// TwinCAT 3 PLC project HalfBROTTests
// Title: HalfBROTTests
// Company: BROT
// ProjectVersion: 0.1.0
// ProgramVersion: 3.1.4024.66
// libraries:
//   HalfBROT, * (BROT)
//   BROTLib, 0.26.0 (BROT)
//   Tc2_Math, * (Beckhoff Automation GmbH)
//   Tc2_MC2, * (Beckhoff Automation GmbH)
//   Tc2_Standard, * (Beckhoff Automation GmbH)
//   Tc2_System, * (Beckhoff Automation GmbH)
//   Tc2_Utilities, * (Beckhoff Automation GmbH)
//   Tc3_Module, * (Beckhoff Automation GmbH)
//   VisuElemEventTable, 1.0.3.0 (System)
//   TcUnit, * (www.tcunit.org)
// project tree:
//   / PlcTask.TcTTO
//   POUs/ F_Note.TcPOU, GVL_Diag.TcGVL, FB_NullComm.TcPOU, FB_TestBase.TcPOU, FB_HydraulicsRig.TcPOU, FB_CoverRig.TcPOU, FB_PendantRig.TcPOU, FB_FocusUnlockRig.TcPOU, FB_HydraulicsControl_Tests.TcPOU, FB_CoverControl_Tests.TcPOU, FB_PendantControl_Tests.TcPOU, FB_FocusUnlock_Tests.TcPOU, FB_BrakeCloseHold_Tests.TcPOU, F_FocusHoldOnStop_Tests.TcPOU, MAIN.TcPOU
// real-time tasks:
//   TASK PlcTask: cycle T#10ms, priority 20, ADS port 350

CONFIGURATION HalfBROTTests
    RESOURCE PLC ON TwinCAT3
        TASK PlcTask(INTERVAL := T#10ms, PRIORITY := 20);
        PROGRAM MAIN WITH PlcTask : MAIN;
    END_RESOURCE
END_CONFIGURATION

// ---- POUs/GVL_Diag.TcGVL
{attribute 'qualified_only'}
VAR_GLOBAL
	// the failed checks of the scenario tests (F_Note), one "test: message;" each. Run-Tests.ps1 prints it when a test failed:
	// TcUnit itself only writes the failure text to the ADS log, which CI cannot see.
	sFailures	: STRING(1000);
END_VAR

// ---- POUs/MAIN.TcPOU
PROGRAM MAIN
VAR
	// TcUnit finds every FB_TestSuite instance by itself; it is enough to declare them here.
	fbHydraulicsTests	: FB_HydraulicsControl_Tests;
	fbCoverTests		: FB_CoverControl_Tests;
	fbPendantTests		: FB_PendantControl_Tests;
	fbFocusUnlockTests	: FB_FocusUnlock_Tests;
	fbBrakeCloseHoldTests	: FB_BrakeCloseHold_Tests;	// MONETcommon#277
	fbFocusHoldOnStopTests	: F_FocusHoldOnStop_Tests;	// MONETcommon#278
END_VAR

TcUnit.RUN();

END_PROGRAM

// ---- POUs/FB_HydraulicsControl_Tests.TcPOU
// Characterisation tests of HalfBROT.FB_HydraulicsControl (HalfBROT#32 step 3) through the I/O structs and the command methods
// (#30, #31): start-up, the brake (pressure delay, clearing, pressure loss, CloseBrake, pump stop, azimuth limit), the manual
// brake re-arm of #31, and the latched errors that need no more than 13 s. They pin what the block does today, they are
// not a specification. Every test owns a rig (FB_HydraulicsRig, a plant behind the structs) and runs over many PLC cycles;
// the block timers run on the system time, so the tests take real time (the longest about 15 s). The suction and
// pressure watchdogs are shortened through tSuctionWatchdog and tPressureWatchdog.
FUNCTION_BLOCK FB_HydraulicsControl_Tests EXTENDS FB_TestBase
VAR
END_VAR

Idle_Everything_Off();
Enable_Runs_Pump();
Open_Brake_After_Pressure_Delay();
No_Clearing_Keeps_Brake_Closed();
Pressure_Loss_Closes_Brake_Auto_Reopens();
CloseBrake_Closes_And_Ends_Request();
Pump_Stop_Closes_Brake();
Azimuth_Limit_Closes_Brake();
Manual_Brake_Stays_Closed_After_Pressure_Loss();
Manual_Brake_Reopens_After_Switch_Off_On();
Manual_Switch_Off_Closes_Brake();
Manual_Brake_Stays_Closed_After_Pump_Restart();
Oil_Low_Is_Error_Until_Reset();
Hydraulics_Watchdog_Is_Error();
Suction_Without_Feedback_Is_Error();
Missing_Pressure_Is_Error();
Main_Pump_Without_Feedback_Is_Error();

// No request, healthy sensors: no pump, no brake, no error, no starter reset.
METHOD PRIVATE Idle_Everything_Off
VAR_INST
	rig		: FB_HydraulicsRig;
	nStep	: INT;
	bViol	: BOOL;
END_VAR
TEST('Idle_Everything_Off');
sCurrent := 'Idle_Everything_Off: ';
IF nStep >= 90 THEN
	RETURN;
END_IF
rig.Scan();
IF rig.nScans >= 5 THEN
	Check(NOT rig.stOut.bOilPumpEnable, 'no pump enable');
	Check(NOT rig.stOut.bOilSuctionEnable, 'no suction enable');
	Check(NOT rig.stOut.bBrakeAzEl, 'brake output off');
	Check(NOT rig.fb.bError, 'no error with healthy sensors');
	Check(rig.fb.PumpState = HalfBROT.E_PumpState.Off, 'pump state Off');
	Check(rig.fb.bBrakeClosed AND NOT rig.fb.bBrakeOpen, 'brake reported closed');
	Check(rig.fb.BrakeState = HalfBROT.E_BrakeState.Closed, 'brake state Closed');
	Check(NOT rig.stOut.bResetOilPump AND NOT rig.stOut.bResetSuctionPump, 'no starter reset');
		nStep := 99;
		TEST_FINISHED();
END_IF
END_METHOD

// Enable starts the pump; the plant reports it running with pressure; the brake is not opened by the pump start.
METHOD PRIVATE Enable_Runs_Pump
VAR_INST
	rig		: FB_HydraulicsRig;
	nStep	: INT;
	bViol	: BOOL;
END_VAR
TEST('Enable_Runs_Pump');
sCurrent := 'Enable_Runs_Pump: ';
IF nStep >= 90 THEN
	RETURN;
END_IF
rig.Scan();
CASE nStep OF
0:
	rig.SetEnable(TRUE);
	rig.StepStart();
	nStep := 10;
10:
	IF rig.nStepScans >= 6 THEN
		Check(rig.fb.Enable, 'Enable reads back');
		Check(rig.stOut.bOilPumpEnable, 'pump enable output');
		Check(rig.fb.PumpRunning AND rig.fb.OilPressureOK, 'pump running and pressure reported');
		Check(rig.fb.PumpState = HalfBROT.E_PumpState.Running, 'pump state Running');
		Check(NOT rig.fb.Error, 'no error');
		Check(NOT rig.stOut.bBrakeAzEl, 'the pump start does not open the brake');
		nStep := 99;
		TEST_FINISHED();
	END_IF
END_CASE
END_METHOD

// OpenBrake() each scan: the brake output comes about 3 s after the pressure, the report 1 s after the output.
METHOD PRIVATE Open_Brake_After_Pressure_Delay
VAR_INST
	rig		: FB_HydraulicsRig;
	nStep	: INT;
	bViol	: BOOL;
END_VAR
TEST('Open_Brake_After_Pressure_Delay');
sCurrent := 'Open_Brake_After_Pressure_Delay: ';
IF nStep >= 90 THEN
	RETURN;
END_IF
rig.Scan();
CASE nStep OF
0:
	rig.bClearing := TRUE;
	rig.bAuto := TRUE;
	rig.SetEnable(TRUE);
	rig.StepStart();
	nStep := 10;
10:
	IF rig.StepTime(T#1S) THEN
		Check(NOT rig.stOut.bBrakeAzEl, 'no brake output during the pressure delay');
		nStep := 20;
	END_IF
20:
	IF rig.stOut.bBrakeAzEl THEN
		Check(rig.StepTime(T#2S500MS) AND NOT rig.StepTime(T#4S), 'the brake output comes about 3 s after the start');
		Check(NOT rig.fb.bBrakeOpen, 'open is reported 1 s after the output, not with it');
		Check(rig.fb.BrakeState = HalfBROT.E_BrakeState.Opening, 'brake state Opening while the output is on and not reported');
		rig.StepStart();
		nStep := 30;
	ELSIF rig.StepTime(T#6S) THEN
		Check(FALSE, 'the brake output never came');
		nStep := 99;
		TEST_FINISHED();
	END_IF
30:
	IF rig.fb.bBrakeOpen THEN
		Check(rig.StepTime(T#800MS) AND NOT rig.StepTime(T#2S), 'open is reported about 1 s after the output');
		Check(rig.fb.BrakeOpen AND NOT rig.fb.bBrakeClosed, 'BrakeOpen property and bBrakeClosed agree');
		Check(rig.fb.BrakeState = HalfBROT.E_BrakeState.Open, 'brake state Open when reported');
		nStep := 99;
		TEST_FINISHED();
	ELSIF rig.StepTime(T#3S) THEN
		Check(FALSE, 'open was never reported');
		nStep := 99;
		TEST_FINISHED();
	END_IF
END_CASE
END_METHOD

// Without bBrakeClearing the brake is not opened although it is requested and the pressure is there.
METHOD PRIVATE No_Clearing_Keeps_Brake_Closed
VAR_INST
	rig		: FB_HydraulicsRig;
	nStep	: INT;
	bViol	: BOOL;
END_VAR
TEST('No_Clearing_Keeps_Brake_Closed');
sCurrent := 'No_Clearing_Keeps_Brake_Closed: ';
IF nStep >= 90 THEN
	RETURN;
END_IF
rig.Scan();
CASE nStep OF
0:
	rig.bClearing := FALSE;
	rig.bAuto := TRUE;
	rig.SetEnable(TRUE);
	rig.StepStart();
	nStep := 10;
10:
	bViol := bViol OR rig.stOut.bBrakeAzEl OR rig.fb.bBrakeOpen;
	IF rig.StepTime(T#4S) THEN
		Check(NOT bViol, 'the brake stays closed without the clearing');
		Check(rig.fb.PumpRunning AND rig.fb.OilPressureOK, 'pump running with pressure');
		nStep := 99;
		TEST_FINISHED();
	END_IF
END_CASE
END_METHOD

// Pressure loss closes the brake after the 2 s debounce; with the automatic request still there it opens again after the pressure delay.
METHOD PRIVATE Pressure_Loss_Closes_Brake_Auto_Reopens
VAR_INST
	rig		: FB_HydraulicsRig;
	nStep	: INT;
	bViol	: BOOL;
END_VAR
TEST('Pressure_Loss_Closes_Brake_Auto_Reopens');
sCurrent := 'Pressure_Loss_Closes_Brake_Auto_Reopens: ';
IF nStep >= 90 THEN
	RETURN;
END_IF
rig.Scan();
CASE nStep OF
0:
	rig.bClearing := TRUE;
	rig.bAuto := TRUE;
	rig.SetEnable(TRUE);
	rig.StepStart();
	nStep := 10;
10:
	IF rig.fb.bBrakeOpen THEN
		rig.bPressure := FALSE;
		rig.StepStart();
		nStep := 20;
	ELSIF rig.StepTime(T#8S) THEN
		Check(FALSE, 'the brake never opened');
		nStep := 99;
		TEST_FINISHED();
	END_IF
20:
	IF NOT rig.stOut.bBrakeAzEl THEN
		Check(rig.StepTime(T#1S500MS), 'the brake holds during the 2 s debounce');
		Check(NOT rig.fb.bBrakeOpen, 'closed is reported');
		Check(rig.stOut.bOilPumpEnable, 'the pump enable stays');
		rig.bPressure := TRUE;
		rig.StepStart();
		nStep := 30;
	ELSIF rig.StepTime(T#4S) THEN
		Check(FALSE, 'the brake did not close on the pressure loss');
		nStep := 99;
		TEST_FINISHED();
	END_IF
30:
	IF rig.stOut.bBrakeAzEl THEN
		Check(rig.StepTime(T#2S), 'the brake opens again only after the pressure delay');
		nStep := 99;
		TEST_FINISHED();
	ELSIF rig.StepTime(T#6S) THEN
		Check(FALSE, 'the automatic request did not open the brake again');
		nStep := 99;
		TEST_FINISHED();
	END_IF
END_CASE
END_METHOD

// CloseBrake() closes the brake at once and the request ends: no automatic re-open without OpenBrake().
METHOD PRIVATE CloseBrake_Closes_And_Ends_Request
VAR_INST
	rig		: FB_HydraulicsRig;
	nStep	: INT;
	bViol	: BOOL;
END_VAR
TEST('CloseBrake_Closes_And_Ends_Request');
sCurrent := 'CloseBrake_Closes_And_Ends_Request: ';
IF nStep >= 90 THEN
	RETURN;
END_IF
rig.Scan();
CASE nStep OF
0:
	rig.bClearing := TRUE;
	rig.bAuto := TRUE;
	rig.SetEnable(TRUE);
	rig.StepStart();
	nStep := 10;
10:
	IF rig.fb.bBrakeOpen THEN
		rig.bAuto := FALSE;
		rig.fb.CloseBrake();
		rig.StepStart();
		nStep := 20;
	ELSIF rig.StepTime(T#8S) THEN
		Check(FALSE, 'the brake never opened');
		nStep := 99;
		TEST_FINISHED();
	END_IF
20:
	IF NOT rig.stOut.bBrakeAzEl THEN
		Check(NOT rig.StepTime(T#300MS), 'the brake output drops at once');
		Check(NOT rig.fb.bBrakeOpen, 'closed is reported');
		Check(rig.fb.BrakeState = HalfBROT.E_BrakeState.Closed, 'brake state Closed after the close');
		rig.StepStart();
		nStep := 30;
	ELSIF rig.StepTime(T#1S) THEN
		Check(FALSE, 'CloseBrake() did not close the brake');
		nStep := 99;
		TEST_FINISHED();
	END_IF
30:
	bViol := bViol OR rig.stOut.bBrakeAzEl;
	IF rig.StepTime(T#4S) THEN
		Check(NOT bViol, 'the brake stays closed with the pressure there');
		nStep := 99;
		TEST_FINISHED();
	END_IF
END_CASE
END_METHOD

// ManualStopPump drops the pump enable; with the pump the brake closes.
METHOD PRIVATE Pump_Stop_Closes_Brake
VAR_INST
	rig		: FB_HydraulicsRig;
	nStep	: INT;
	bViol	: BOOL;
END_VAR
TEST('Pump_Stop_Closes_Brake');
sCurrent := 'Pump_Stop_Closes_Brake: ';
IF nStep >= 90 THEN
	RETURN;
END_IF
rig.Scan();
CASE nStep OF
0:
	rig.bClearing := TRUE;
	rig.bAuto := TRUE;
	rig.SetEnable(TRUE);
	rig.StepStart();
	nStep := 10;
10:
	IF rig.fb.bBrakeOpen THEN
		rig.bAuto := FALSE;
		rig.SetStopPump(TRUE);
		rig.StepStart();
		nStep := 20;
	ELSIF rig.StepTime(T#8S) THEN
		Check(FALSE, 'the brake never opened');
		nStep := 99;
		TEST_FINISHED();
	END_IF
20:
	IF NOT rig.stOut.bBrakeAzEl THEN
		Check(NOT rig.StepTime(T#300MS), 'the brake output drops with the pump');
		Check(NOT rig.stOut.bOilPumpEnable, 'pump enable off');
		Check(NOT rig.fb.bBrakeOpen, 'closed is reported');
		nStep := 99;
		TEST_FINISHED();
	ELSIF rig.StepTime(T#1S) THEN
		Check(FALSE, 'the pump stop did not close the brake');
		nStep := 99;
		TEST_FINISHED();
	END_IF
END_CASE
END_METHOD

// The azimuth limit switch closes the brake and holds it closed while it is active, although the request goes on.
METHOD PRIVATE Azimuth_Limit_Closes_Brake
VAR_INST
	rig		: FB_HydraulicsRig;
	nStep	: INT;
	bViol	: BOOL;
END_VAR
TEST('Azimuth_Limit_Closes_Brake');
sCurrent := 'Azimuth_Limit_Closes_Brake: ';
IF nStep >= 90 THEN
	RETURN;
END_IF
rig.Scan();
CASE nStep OF
0:
	rig.bClearing := TRUE;
	rig.bAuto := TRUE;
	rig.SetEnable(TRUE);
	rig.StepStart();
	nStep := 10;
10:
	IF rig.fb.bBrakeOpen THEN
		rig.bAzLimit := TRUE;
		rig.StepStart();
		nStep := 20;
	ELSIF rig.StepTime(T#8S) THEN
		Check(FALSE, 'the brake never opened');
		nStep := 99;
		TEST_FINISHED();
	END_IF
20:
	IF NOT rig.stOut.bBrakeAzEl THEN
		Check(NOT rig.StepTime(T#300MS), 'the brake output drops at once');
		rig.StepStart();
		nStep := 30;
	ELSIF rig.StepTime(T#1S) THEN
		Check(FALSE, 'the azimuth limit did not close the brake');
		nStep := 99;
		TEST_FINISHED();
	END_IF
30:
	bViol := bViol OR rig.stOut.bBrakeAzEl;
	IF rig.StepTime(T#4S) THEN
		Check(NOT bViol, 'the brake stays closed while the limit is active');
		nStep := 99;
		TEST_FINISHED();
	END_IF
END_CASE
END_METHOD

// #31: the cabinet switch opens the brake once; after a pressure loss it stays closed while the switch stays on, with the pressure back.
METHOD PRIVATE Manual_Brake_Stays_Closed_After_Pressure_Loss
VAR_INST
	rig		: FB_HydraulicsRig;
	nStep	: INT;
	bViol	: BOOL;
END_VAR
TEST('Manual_Brake_Stays_Closed_After_Pressure_Loss');
sCurrent := 'Manual_Brake_Stays_Closed_After_Pressure_Loss: ';
IF nStep >= 90 THEN
	RETURN;
END_IF
rig.Scan();
CASE nStep OF
0:
	// the pump runs first: a switch edge before the pump runs is dropped by the block (the request is cleared while the pump is off)
	rig.bManual := TRUE;
	rig.SetEnable(TRUE);
	rig.StepStart();
	nStep := 5;
5:
	IF rig.StepTime(T#500MS) THEN
		rig.bSwitch := TRUE;
		rig.StepStart();
		nStep := 10;
	END_IF
10:
	IF rig.fb.bBrakeOpen THEN
		Check(rig.stOut.bBrakeAzEl, 'the switch opened the brake');
		rig.bPressure := FALSE;
		rig.StepStart();
		nStep := 20;
	ELSIF rig.StepTime(T#8S) THEN
		Check(FALSE, 'the brake never opened');
		nStep := 99;
		TEST_FINISHED();
	END_IF
20:
	IF NOT rig.stOut.bBrakeAzEl THEN
		Check(rig.StepTime(T#1S500MS), 'the brake holds during the 2 s debounce');
		rig.bPressure := TRUE;
		bViol := FALSE;
		rig.StepStart();
		nStep := 30;
	ELSIF rig.StepTime(T#4S) THEN
		Check(FALSE, 'the brake did not close on the pressure loss');
		nStep := 99;
		TEST_FINISHED();
	END_IF
30:
	bViol := bViol OR rig.stOut.bBrakeAzEl;
	IF rig.StepTime(T#4S500MS) THEN
		Check(rig.fb.bOilPressureOK AND rig.fb.PumpRunning, 'pressure is back');
		Check(NOT bViol, 'the brake is not opened again while the switch stays on');
		nStep := 99;
		TEST_FINISHED();
	END_IF
END_CASE
END_METHOD

// #31: after CloseBrake() the brake stays closed while the switch stays on; switch off and on opens it again.
METHOD PRIVATE Manual_Brake_Reopens_After_Switch_Off_On
VAR_INST
	rig		: FB_HydraulicsRig;
	nStep	: INT;
	bViol	: BOOL;
END_VAR
TEST('Manual_Brake_Reopens_After_Switch_Off_On');
sCurrent := 'Manual_Brake_Reopens_After_Switch_Off_On: ';
IF nStep >= 90 THEN
	RETURN;
END_IF
rig.Scan();
CASE nStep OF
0:
	// the pump runs first: a switch edge before the pump runs is dropped by the block (the request is cleared while the pump is off)
	rig.bManual := TRUE;
	rig.SetEnable(TRUE);
	rig.StepStart();
	nStep := 5;
5:
	IF rig.StepTime(T#500MS) THEN
		rig.bSwitch := TRUE;
		rig.StepStart();
		nStep := 10;
	END_IF
10:
	IF rig.fb.bBrakeOpen THEN
		rig.fb.CloseBrake();
		rig.StepStart();
		nStep := 20;
	ELSIF rig.StepTime(T#8S) THEN
		Check(FALSE, 'the brake never opened');
		nStep := 99;
		TEST_FINISHED();
	END_IF
20:
	IF NOT rig.stOut.bBrakeAzEl THEN
		Check(NOT rig.StepTime(T#300MS), 'CloseBrake() closes at once');
		bViol := FALSE;
		rig.StepStart();
		nStep := 30;
	ELSIF rig.StepTime(T#1S) THEN
		Check(FALSE, 'CloseBrake() did not close the brake');
		nStep := 99;
		TEST_FINISHED();
	END_IF
30:
	bViol := bViol OR rig.stOut.bBrakeAzEl;
	IF rig.StepTime(T#4S) THEN
		Check(NOT bViol, 'the brake stays closed while the switch stays on');
		rig.bSwitch := FALSE;
		rig.StepStart();
		nStep := 40;
	END_IF
40:
	IF rig.StepTime(T#500MS) THEN
		Check(NOT rig.stOut.bBrakeAzEl, 'the brake is closed with the switch off');
		rig.bSwitch := TRUE;
		rig.StepStart();
		nStep := 50;
	END_IF
50:
	IF rig.stOut.bBrakeAzEl THEN
		Check(NOT rig.StepTime(T#1S), 'the switch off and on opens the brake at once, the pressure delay has long run out');
		nStep := 99;
		TEST_FINISHED();
	ELSIF rig.StepTime(T#6S) THEN
		Check(FALSE, 'the brake did not open again after the switch went off and on');
		nStep := 99;
		TEST_FINISHED();
	END_IF
END_CASE
END_METHOD

// The permission: switch off closes the brake at once (bBrakeClearing) and ends the request.
METHOD PRIVATE Manual_Switch_Off_Closes_Brake
VAR_INST
	rig		: FB_HydraulicsRig;
	nStep	: INT;
	bViol	: BOOL;
END_VAR
TEST('Manual_Switch_Off_Closes_Brake');
sCurrent := 'Manual_Switch_Off_Closes_Brake: ';
IF nStep >= 90 THEN
	RETURN;
END_IF
rig.Scan();
CASE nStep OF
0:
	// the pump runs first: a switch edge before the pump runs is dropped by the block (the request is cleared while the pump is off)
	rig.bManual := TRUE;
	rig.SetEnable(TRUE);
	rig.StepStart();
	nStep := 5;
5:
	IF rig.StepTime(T#500MS) THEN
		rig.bSwitch := TRUE;
		rig.StepStart();
		nStep := 10;
	END_IF
10:
	IF rig.fb.bBrakeOpen THEN
		rig.bSwitch := FALSE;
		rig.StepStart();
		nStep := 20;
	ELSIF rig.StepTime(T#8S) THEN
		Check(FALSE, 'the brake never opened');
		nStep := 99;
		TEST_FINISHED();
	END_IF
20:
	IF NOT rig.stOut.bBrakeAzEl THEN
		Check(NOT rig.StepTime(T#300MS), 'the brake output drops at once');
		Check(NOT rig.fb.bBrakeOpen, 'closed is reported');
		Check(rig.fb.BrakeState = HalfBROT.E_BrakeState.Closed, 'brake state Closed after the close');
		nStep := 99;
		TEST_FINISHED();
	ELSIF rig.StepTime(T#1S) THEN
		Check(FALSE, 'the switch off did not close the brake');
		nStep := 99;
		TEST_FINISHED();
	END_IF
END_CASE
END_METHOD

// #31: a pump stop closes the brake; the pump runs again with the switch still on: the brake stays closed.
METHOD PRIVATE Manual_Brake_Stays_Closed_After_Pump_Restart
VAR_INST
	rig		: FB_HydraulicsRig;
	nStep	: INT;
	bViol	: BOOL;
END_VAR
TEST('Manual_Brake_Stays_Closed_After_Pump_Restart');
sCurrent := 'Manual_Brake_Stays_Closed_After_Pump_Restart: ';
IF nStep >= 90 THEN
	RETURN;
END_IF
rig.Scan();
CASE nStep OF
0:
	// the pump runs first: a switch edge before the pump runs is dropped by the block (the request is cleared while the pump is off)
	rig.bManual := TRUE;
	rig.SetEnable(TRUE);
	rig.StepStart();
	nStep := 5;
5:
	IF rig.StepTime(T#500MS) THEN
		rig.bSwitch := TRUE;
		rig.StepStart();
		nStep := 10;
	END_IF
10:
	IF rig.fb.bBrakeOpen THEN
		rig.SetStopPump(TRUE);
		rig.StepStart();
		nStep := 20;
	ELSIF rig.StepTime(T#8S) THEN
		Check(FALSE, 'the brake never opened');
		nStep := 99;
		TEST_FINISHED();
	END_IF
20:
	IF NOT rig.stOut.bBrakeAzEl THEN
		Check(NOT rig.StepTime(T#300MS), 'the pump stop closes the brake at once');
		rig.StepStart();
		nStep := 30;
	ELSIF rig.StepTime(T#1S) THEN
		Check(FALSE, 'the pump stop did not close the brake');
		nStep := 99;
		TEST_FINISHED();
	END_IF
30:
	IF rig.StepTime(T#500MS) THEN
		rig.SetStopPump(FALSE);
		bViol := FALSE;
		rig.StepStart();
		nStep := 40;
	END_IF
40:
	bViol := bViol OR rig.stOut.bBrakeAzEl;
	IF rig.StepTime(T#4S500MS) THEN
		Check(rig.fb.PumpRunning AND rig.fb.OilPressureOK, 'the pump runs again with pressure');
		Check(NOT bViol, 'the brake is not opened again while the switch stays on');
		nStep := 99;
		TEST_FINISHED();
	END_IF
END_CASE
END_METHOD

// Oil low is a latched error that stops the pump; Reset() clears it once the oil is back and the pump starts again (Enable is still set).
METHOD PRIVATE Oil_Low_Is_Error_Until_Reset
VAR_INST
	rig		: FB_HydraulicsRig;
	nStep	: INT;
	bViol	: BOOL;
END_VAR
TEST('Oil_Low_Is_Error_Until_Reset');
sCurrent := 'Oil_Low_Is_Error_Until_Reset: ';
IF nStep >= 90 THEN
	RETURN;
END_IF
rig.Scan();
CASE nStep OF
0:
	rig.SetEnable(TRUE);
	rig.StepStart();
	nStep := 10;
10:
	IF rig.nStepScans >= 5 THEN
		rig.stIn.bOilLow := FALSE;
		rig.StepStart();
		nStep := 20;
	END_IF
20:
	IF rig.nStepScans >= 3 THEN
		Check(rig.fb.Error AND rig.fb.bOilLow, 'oil low is an error');
		Check(rig.fb.PumpState = HalfBROT.E_PumpState.Error, 'pump state Error');
		Check(NOT rig.stOut.bOilPumpEnable, 'the error stops the pump');
		rig.stIn.bOilLow := TRUE;
		rig.StepStart();
		nStep := 30;
	END_IF
30:
	IF rig.nStepScans >= 3 THEN
		Check(rig.fb.Error, 'the error stays latched with the oil back');
		rig.fb.Reset();
		rig.StepStart();
		nStep := 40;
	END_IF
40:
	IF rig.nStepScans >= 4 THEN
		Check(NOT rig.fb.Error, 'Reset() clears the error');
		Check(rig.stOut.bOilPumpEnable, 'the pump starts again, Enable is still set');
		Check(rig.fb.PumpState = HalfBROT.E_PumpState.Running, 'pump state Running again after Reset()');
		nStep := 99;
		TEST_FINISHED();
	END_IF
END_CASE
END_METHOD

// The pump running without the suction pump for tHydraulicsWatchdog (1 s here, 140 s default, #10) is a latched error.
METHOD PRIVATE Hydraulics_Watchdog_Is_Error
VAR_INST
	rig		: FB_HydraulicsRig;
	nStep	: INT;
	bViol	: BOOL;
END_VAR
TEST('Hydraulics_Watchdog_Is_Error');
sCurrent := 'Hydraulics_Watchdog_Is_Error: ';
IF nStep >= 90 THEN
	RETURN;
END_IF
rig.Scan();
CASE nStep OF
0:
	rig.tHydraulicsWatchdog := T#1S;
	rig.bSuctionFollows := FALSE;
	rig.SetEnable(TRUE);
	rig.StepStart();
	nStep := 10;
10:
	bViol := bViol OR rig.fb.bHydraulicsFailure;
	IF rig.fb.Error THEN
		Check(rig.StepTime(T#800MS), 'not before the configured time');
		Check(bViol, 'the hydraulics failure was reported');
		Check(NOT rig.stOut.bOilPumpEnable, 'the error stops the pump');
		nStep := 99;
		TEST_FINISHED();
	ELSIF rig.StepTime(T#4S) THEN
		Check(FALSE, 'no hydraulics failure');
		nStep := 99;
		TEST_FINISHED();
	END_IF
END_CASE
END_METHOD

// The suction enable (manual start) without the run feedback for tSuctionWatchdog (1 s here, 15 s default) is a latched error.
METHOD PRIVATE Suction_Without_Feedback_Is_Error
VAR_INST
	rig		: FB_HydraulicsRig;
	nStep	: INT;
	bViol	: BOOL;
END_VAR
TEST('Suction_Without_Feedback_Is_Error');
sCurrent := 'Suction_Without_Feedback_Is_Error: ';
IF nStep >= 90 THEN
	RETURN;
END_IF
rig.Scan();
CASE nStep OF
0:
	rig.tSuctionWatchdog := T#1S;
	rig.bSuctionFollows := FALSE;
	rig.SetSuction(TRUE);
	rig.StepStart();
	nStep := 10;
10:
	bViol := bViol OR rig.fb.bSuctionFailure;
	IF rig.fb.Error THEN
		Check(rig.stOut.bOilSuctionEnable, 'the suction enable was on');
		Check(rig.StepTime(T#800MS), 'not before the configured time');
		Check(bViol, 'the suction failure was reported');
		nStep := 99;
		TEST_FINISHED();
	ELSIF rig.StepTime(T#4S) THEN
		Check(FALSE, 'no suction failure');
		nStep := 99;
		TEST_FINISHED();
	END_IF
END_CASE
END_METHOD

// The pump enabled without oil pressure for tPressureWatchdog (1 s here, 30 s default) is a latched error that stops the pump.
METHOD PRIVATE Missing_Pressure_Is_Error
VAR_INST
	rig		: FB_HydraulicsRig;
	nStep	: INT;
	bViol	: BOOL;
END_VAR
TEST('Missing_Pressure_Is_Error');
sCurrent := 'Missing_Pressure_Is_Error: ';
IF nStep >= 90 THEN
	RETURN;
END_IF
rig.Scan();
CASE nStep OF
0:
	rig.tPressureWatchdog := T#1S;
	rig.bPressure := FALSE;
	rig.SetEnable(TRUE);
	rig.StepStart();
	nStep := 10;
10:
	bViol := bViol OR rig.fb.bPressureFailure;
	IF rig.fb.Error THEN
		Check(rig.StepTime(T#800MS), 'not before the configured time');
		Check(bViol, 'the pressure failure was reported');
		Check(NOT rig.stOut.bOilPumpEnable, 'the error stops the pump');
		nStep := 99;
		TEST_FINISHED();
	ELSIF rig.StepTime(T#4S) THEN
		Check(FALSE, 'no pressure failure');
		nStep := 99;
		TEST_FINISHED();
	END_IF
END_CASE
END_METHOD

// No run feedback 10 s after the pump enable is a latched error (main pump failure).
METHOD PRIVATE Main_Pump_Without_Feedback_Is_Error
VAR_INST
	rig		: FB_HydraulicsRig;
	nStep	: INT;
	bViol	: BOOL;
END_VAR
TEST('Main_Pump_Without_Feedback_Is_Error');
sCurrent := 'Main_Pump_Without_Feedback_Is_Error: ';
IF nStep >= 90 THEN
	RETURN;
END_IF
rig.Scan();
CASE nStep OF
0:
	rig.bPumpFollows := FALSE;
	rig.SetEnable(TRUE);
	rig.StepStart();
	nStep := 10;
10:
	bViol := bViol OR rig.fb.bMainPumpFailure;
	IF rig.fb.Error THEN
		Check(rig.StepTime(T#9S500MS), 'not before the 10 s');
		Check(bViol, 'the main pump failure was reported');
		Check(NOT rig.stOut.bOilPumpEnable, 'the error stops the pump');
		nStep := 99;
		TEST_FINISHED();
	ELSIF rig.StepTime(T#13S) THEN
		Check(FALSE, 'no main pump failure');
		nStep := 99;
		TEST_FINISHED();
	END_IF
END_CASE
END_METHOD

END_FUNCTION_BLOCK

// ---- POUs/FB_TestBase.TcPOU
// Base of the HalfBROTTests suites: Check() is a TcUnit assertion that also notes a failed check in GVL_Diag.sFailures
// (printed by tools/Run-Tests.ps1, TcUnit itself writes the failure text only to the ADS log). The test method sets
// sCurrent to its name first.
FUNCTION_BLOCK FB_TestBase EXTENDS TcUnit.FB_TestSuite
VAR
	sCurrent	: STRING(80);
END_VAR

METHOD Check
VAR_INPUT
	bCondition	: BOOL;
	sMessage	: STRING(255);
END_VAR
AssertTrue(Condition := bCondition, Message := sMessage);
F_Note(bFailed := NOT bCondition, sText := CONCAT(sCurrent, sMessage));
END_METHOD

END_FUNCTION_BLOCK

// ---- POUs/F_Note.TcPOU
// Records a failed check in GVL_Diag.sFailures (see there). Called next to the TcUnit assertion, which does the actual test result.
FUNCTION F_Note : BOOL
VAR_INPUT
	bFailed	: BOOL;
	sText	: STRING(255);
END_VAR

IF bFailed AND LEN(GVL_Diag.sFailures) < 700 THEN
	GVL_Diag.sFailures := CONCAT(CONCAT(GVL_Diag.sFailures, sText), '; ');
END_IF
F_Note := bFailed;

END_FUNCTION

// ---- POUs/FB_HydraulicsRig.TcPOU
// FB_HydraulicsControl with a plant: the pump feedback follows the pump enable output one scan later and the oil pressure
// follows the pump (a starter and a pump that work), the suction feedback follows the suction enable. The sensors are healthy.
// bAuto calls OpenBrake() in every scan (the automatic request of MONETcommon), bManual calls ManualBrake(bSwitch) and
// feeds the switch to bBrakeClearing as MAIN of MONETS/MONETN does. tPumpResetPulse is T#0S: the pump starts at once.
// StepStart()/StepTime() measure real time from the start of a step (the block timers run on the system time).
FUNCTION_BLOCK FB_HydraulicsRig
VAR_INPUT
	stIn		: HalfBROT.ST_HydraulicsIn := (bOilLow := TRUE, bOilHigh := TRUE, bOilCold := TRUE, bOilFilterDirty := TRUE, nOilLevel := 8000);
	bClearing	: BOOL;
	bAzLimit	: BOOL;
	bAuto		: BOOL;
	bManual		: BOOL;
	bSwitch		: BOOL;
	bPumpFollows	: BOOL := TRUE;
	bPressure		: BOOL := TRUE;
	bSuctionFollows	: BOOL := TRUE;
	tHydraulicsWatchdog	: TIME := T#140S;
	tSuctionWatchdog	: TIME := T#15S;
	tPressureWatchdog	: TIME := T#30S;
END_VAR
VAR
	fbComm		: FB_NullComm;
	fb			: HalfBROT.FB_HydraulicsControl(comm := fbComm);
	stOut		: HalfBROT.ST_HydraulicsOut;
	tonStep		: TON;
	nScans		: UDINT;
	nStepScans	: UDINT;
END_VAR

METHOD Scan
nScans := nScans + 1;
nStepScans := nStepScans + 1;
IF bPumpFollows THEN
	stIn.bPumpRunning := stOut.bOilPumpEnable;
END_IF
stIn.bOilPressureOK := stIn.bPumpRunning AND bPressure;
IF bSuctionFollows THEN
	stIn.bSuctionRunning := stOut.bOilSuctionEnable;
END_IF
IF bAuto THEN
	fb.OpenBrake();
END_IF
IF bManual THEN
	bClearing := bSwitch;
	fb.ManualBrake(bSwitch := bSwitch);
END_IF
fb(stIn := stIn, bBrakeClearing := bClearing, bAzimuthLimitSwitch := bAzLimit, tHydraulicsWatchdog := tHydraulicsWatchdog,
	tSuctionWatchdog := tSuctionWatchdog, tPressureWatchdog := tPressureWatchdog, tPumpResetPulse := T#0S, stOut := stOut);
tonStep(IN := TRUE, PT := T#1H);
END_METHOD

METHOD StepStart
tonStep(IN := FALSE, PT := T#1H);
nStepScans := 0;
END_METHOD

METHOD StepTime : BOOL
VAR_INPUT
	tTime	: TIME;
END_VAR
StepTime := tonStep.ET >= tTime;
END_METHOD

METHOD SetEnable
VAR_INPUT
	bOn	: BOOL;
END_VAR
fb.Enable := bOn;
END_METHOD

METHOD SetSuction
VAR_INPUT
	bOn	: BOOL;
END_VAR
fb.ManualStartSuction := bOn;
END_METHOD

METHOD SetStopPump
VAR_INPUT
	bOn	: BOOL;
END_VAR
fb.ManualStopPump := bOn;
END_METHOD

END_FUNCTION_BLOCK

// ---- POUs/FB_NullComm.TcPOU
// Minimal I_Comm stub for tests: every Publish/PublishLog call is a no-op that reports success,
// so FBs under test can call fbComm.Publish(...) freely without a real MQTT connection.
FUNCTION_BLOCK FB_NullComm IMPLEMENTS BROTLib.I_Comm
VAR
END_VAR

METHOD Publish : BOOL
VAR_INPUT
	domain			: STRING(255) := 'environment';
	location		: STRING(255) := 'roof';
	parameter		: STRING(255);
	value			: STRING(255);
END_VAR
VAR_OUTPUT
	published	: BOOL;
END_VAR
Publish := TRUE;
published := TRUE;
END_METHOD

METHOD PublishLREAL : BOOL
VAR_INPUT
	domain			: STRING(255) := 'environment';
	location		: STRING(255) := 'roof';
	parameter		: STRING(255);
	value			: LREAL;
END_VAR
VAR_OUTPUT
	published	: BOOL;
END_VAR
PublishLREAL := TRUE;
published := TRUE;
END_METHOD

METHOD PublishINT : BOOL
VAR_INPUT
	domain			: STRING(255) := 'environment';
	location		: STRING(255) := 'roof';
	parameter		: STRING(255);
	value			: LINT;
END_VAR
VAR_OUTPUT
	published	: BOOL;
END_VAR
PublishINT := TRUE;
published := TRUE;
END_METHOD

METHOD PublishBOOL : BOOL
VAR_INPUT
	domain			: STRING(255) := 'environment';
	location		: STRING(255) := 'roof';
	parameter		: STRING(255);
	value			: BOOL;
END_VAR
VAR_OUTPUT
	published	: BOOL;
END_VAR
PublishBOOL := TRUE;
published := TRUE;
END_METHOD

METHOD PublishString : BOOL
VAR_INPUT
	domain			: STRING(255) := 'environment';
	location		: STRING(255) := 'roof';
	parameter		: STRING(255);
	value			: STRING(255);
END_VAR
VAR_OUTPUT
	published	: BOOL;
END_VAR
PublishString := TRUE;
published := TRUE;
END_METHOD

METHOD PublishLog : BOOL
VAR_INPUT
	level		: STRING(255) := 'INFO';
	message		: STRING(255);
END_VAR
VAR_OUTPUT
	published	: BOOL;
END_VAR
PublishLog := TRUE;
published := TRUE;
END_METHOD

END_FUNCTION_BLOCK

// ---- POUs/FB_CoverControl_Tests.TcPOU
// Characterisation tests of HalfBROT.FB_CoverControl (HalfBROT#32 step 3) through the I/O structs: the sequence 1->3->2 and
// 2->3->1, the last call of Open()/Close() wins, Stop(), the latched error of a limit switch fault (#28), the move timeout and
// the reversal dead time (#27). They pin what the block does today, they are not a specification. Every test owns a rig
// (FB_CoverRig, the limit switches set by hand) and runs over several PLC cycles; the timeout and reversal tests take real time.
FUNCTION_BLOCK FB_CoverControl_Tests EXTENDS FB_TestBase
VAR
END_VAR

Open_Sequence_1_3_2();
Close_Sequence_2_3_1();
Last_Call_Wins_Open_After_Close();
Last_Call_Wins_Close_After_Open();
Stop_Drops_Outputs_And_Command();
Limit_Switch_Fault_Stops_All_Until_Reset();
Move_Timeout_Is_Error();
Reversal_Waits_Dead_Time();

// Open(): cover 1 starts, cover 3 only when 1 is at its open switch, cover 2 only when 1 and 3 are; then all outputs are off.
METHOD PRIVATE Open_Sequence_1_3_2
VAR_INST
	rig		: FB_CoverRig;
	nStep	: INT;
	bViol	: BOOL;
END_VAR
TEST('Open_Sequence_1_3_2');
sCurrent := 'Open_Sequence_1_3_2: ';
IF nStep >= 90 THEN
	RETURN;
END_IF
rig.Scan();
CASE nStep OF
0:
	Check(rig.OpenOutputs() = '---' AND rig.CloseOutputs() = '---', CONCAT('no output without a command ', rig.State()));
	rig.fb.Open();
	nStep := 10;
10:
	Check(rig.OpenOutputs() = 'x--' AND rig.CloseOutputs() = '---', CONCAT('only cover 1 starts ', rig.State()));
	Check(rig.fb.State = HalfBROT.E_CoverState.Opening, CONCAT('state Opening ', rig.State()));
	rig.SetMid(1);
	nStep := 15;
15:
	Check(rig.OpenOutputs() = 'x--', CONCAT('cover 3 waits while cover 1 is on its way ', rig.State()));
	rig.SetOpen(1);
	nStep := 20;
20:
	Check(rig.OpenOutputs() = '--x', CONCAT('cover 3 starts when cover 1 is open ', rig.State()));
	rig.SetMid(3);
	nStep := 25;
25:
	Check(rig.OpenOutputs() = '--x', CONCAT('cover 2 waits while cover 3 is on its way ', rig.State()));
	rig.SetOpen(3);
	nStep := 30;
30:
	Check(rig.OpenOutputs() = '-x-', CONCAT('cover 2 starts when 1 and 3 are open ', rig.State()));
	rig.SetOpen(2);
	nStep := 40;
40:
	Check(rig.fb.bAllOpen AND rig.fb.Opened AND NOT rig.fb.Closed, CONCAT('all covers open ', rig.State()));
	Check(rig.fb.State = HalfBROT.E_CoverState.Idle, CONCAT('state Idle after the last cover ', rig.State()));
	Check(rig.OpenOutputs() = '---' AND rig.CloseOutputs() = '---', CONCAT('all outputs off ', rig.State()));
	nStep := 50;
50:
	Check(rig.OpenOutputs() = '---', CONCAT('the command ended with the last cover ', rig.State()));
	nStep := 99;
	TEST_FINISHED();
END_CASE
END_METHOD

// Close(): cover 2 starts, cover 3 only when 2 is at its closed switch, cover 1 only when 2 and 3 are; then all outputs are off.
METHOD PRIVATE Close_Sequence_2_3_1
VAR_INST
	rig		: FB_CoverRig;
	nStep	: INT;
	bViol	: BOOL;
END_VAR
TEST('Close_Sequence_2_3_1');
sCurrent := 'Close_Sequence_2_3_1: ';
IF nStep >= 90 THEN
	RETURN;
END_IF
rig.Scan();
CASE nStep OF
0:
	rig.AllOpen();
	nStep := 5;
5:
	Check(rig.OpenOutputs() = '---' AND rig.CloseOutputs() = '---', CONCAT('no output without a command ', rig.State()));
	rig.fb.Close();
	nStep := 10;
10:
	Check(rig.CloseOutputs() = '-x-' AND rig.OpenOutputs() = '---', CONCAT('only cover 2 starts ', rig.State()));
	Check(rig.fb.State = HalfBROT.E_CoverState.Closing, CONCAT('state Closing ', rig.State()));
	rig.SetMid(2);
	nStep := 15;
15:
	Check(rig.CloseOutputs() = '-x-', CONCAT('cover 3 waits while cover 2 is on its way ', rig.State()));
	rig.SetClosed(2);
	nStep := 20;
20:
	Check(rig.CloseOutputs() = '--x', CONCAT('cover 3 starts when cover 2 is closed ', rig.State()));
	rig.SetMid(3);
	nStep := 25;
25:
	Check(rig.CloseOutputs() = '--x', CONCAT('cover 1 waits while cover 3 is on its way ', rig.State()));
	rig.SetClosed(3);
	nStep := 30;
30:
	Check(rig.CloseOutputs() = 'x--', CONCAT('cover 1 starts when 2 and 3 are closed ', rig.State()));
	rig.SetClosed(1);
	nStep := 40;
40:
	Check(rig.fb.bAllClosed AND rig.fb.Closed AND NOT rig.fb.Opened, CONCAT('all covers closed ', rig.State()));
	Check(rig.OpenOutputs() = '---' AND rig.CloseOutputs() = '---', CONCAT('all outputs off ', rig.State()));
	nStep := 50;
50:
	Check(rig.CloseOutputs() = '---', CONCAT('the command ended with the last cover ', rig.State()));
	nStep := 99;
	TEST_FINISHED();
END_CASE
END_METHOD

// Close() then Open() in one cycle: the open request wins (Open() drops the close request).
METHOD PRIVATE Last_Call_Wins_Open_After_Close
VAR_INST
	rig		: FB_CoverRig;
	nStep	: INT;
	bViol	: BOOL;
END_VAR
TEST('Last_Call_Wins_Open_After_Close');
sCurrent := 'Last_Call_Wins_Open_After_Close: ';
IF nStep >= 90 THEN
	RETURN;
END_IF
rig.Scan();
CASE nStep OF
0:
	rig.AllMid();
	rig.fb.Close();
	rig.fb.Open();
	nStep := 10;
10:
	Check(rig.CloseOutputs() = '---', CONCAT('no close output ', rig.State()));
	Check(rig.OpenOutputs() = 'x--', CONCAT('cover 1 opens ', rig.State()));
	nStep := 99;
	TEST_FINISHED();
END_CASE
END_METHOD

// Open() then Close() in one cycle: the close request wins (Close() drops the open request).
METHOD PRIVATE Last_Call_Wins_Close_After_Open
VAR_INST
	rig		: FB_CoverRig;
	nStep	: INT;
	bViol	: BOOL;
END_VAR
TEST('Last_Call_Wins_Close_After_Open');
sCurrent := 'Last_Call_Wins_Close_After_Open: ';
IF nStep >= 90 THEN
	RETURN;
END_IF
rig.Scan();
CASE nStep OF
0:
	rig.AllMid();
	rig.fb.Open();
	rig.fb.Close();
	nStep := 10;
10:
	Check(rig.OpenOutputs() = '---', CONCAT('no open output ', rig.State()));
	Check(rig.CloseOutputs() = '-x-', CONCAT('cover 2 closes ', rig.State()));
	nStep := 99;
	TEST_FINISHED();
END_CASE
END_METHOD

// Stop() drops the running output in the next scan and the command with it: nothing restarts.
METHOD PRIVATE Stop_Drops_Outputs_And_Command
VAR_INST
	rig		: FB_CoverRig;
	nStep	: INT;
	bViol	: BOOL;
END_VAR
TEST('Stop_Drops_Outputs_And_Command');
sCurrent := 'Stop_Drops_Outputs_And_Command: ';
IF nStep >= 90 THEN
	RETURN;
END_IF
rig.Scan();
CASE nStep OF
0:
	rig.fb.Open();
	nStep := 10;
10:
	Check(rig.OpenOutputs() = 'x--', CONCAT('cover 1 opens ', rig.State()));
	rig.fb.Stop();
	nStep := 20;
20:
	Check(rig.OpenOutputs() = '---' AND rig.CloseOutputs() = '---', CONCAT('the outputs are off after Stop() ', rig.State()));
	nStep := 30;
30:
	Check(rig.OpenOutputs() = '---', CONCAT('nothing restarts ', rig.State()));
	nStep := 40;
40:
	Check(rig.OpenOutputs() = '---' AND NOT rig.fb.Error, CONCAT('still off, no error ', rig.State()));
	nStep := 99;
	TEST_FINISHED();
END_CASE
END_METHOD

// Both switches of one cover (#28): the error stops all covers and drops the command; it stays latched until Reset(), and the move needs a new Open() after it.
METHOD PRIVATE Limit_Switch_Fault_Stops_All_Until_Reset
VAR_INST
	rig		: FB_CoverRig;
	nStep	: INT;
	bViol	: BOOL;
END_VAR
TEST('Limit_Switch_Fault_Stops_All_Until_Reset');
sCurrent := 'Limit_Switch_Fault_Stops_All_Until_Reset: ';
IF nStep >= 90 THEN
	RETURN;
END_IF
rig.Scan();
CASE nStep OF
0:
	rig.fb.Open();
	nStep := 10;
10:
	Check(rig.OpenOutputs() = 'x--', CONCAT('cover 1 opens ', rig.State()));
	rig.SetBoth(3);
	nStep := 20;
20:
	Check(rig.fb.Error AND rig.fb.bError, CONCAT('the fault is an error ', rig.State()));
	Check(rig.fb.State = HalfBROT.E_CoverState.Error, CONCAT('state Error ', rig.State()));
	Check(rig.OpenOutputs() = '---' AND rig.CloseOutputs() = '---', CONCAT('all covers stop, also those without the fault ', rig.State()));
	rig.SetClosed(3);
	rig.fb.Open();
	nStep := 30;
30:
	Check(rig.fb.Error, CONCAT('the error stays latched with the switch fixed ', rig.State()));
	Check(rig.fb.State = HalfBROT.E_CoverState.Error, CONCAT('state stays Error until Reset() ', rig.State()));
	Check(rig.OpenOutputs() = '---', CONCAT('no output while the error is latched ', rig.State()));
	rig.fb.Reset();
	nStep := 40;
40:
	Check(NOT rig.fb.Error, CONCAT('Reset() clears the error ', rig.State()));
	Check(rig.fb.State = HalfBROT.E_CoverState.Idle, CONCAT('state Idle after Reset() ', rig.State()));
	Check(rig.OpenOutputs() = '---', CONCAT('the command was dropped by the error: nothing moves ', rig.State()));
	rig.fb.Open();
	nStep := 50;
50:
	Check(rig.OpenOutputs() = 'x--', CONCAT('a new Open() moves again ', rig.State()));
	nStep := 99;
	TEST_FINISHED();
END_CASE
END_METHOD

// A cover driven for tMoveTimeout (300 ms here, 60 s default) without reaching its switch stops and latches an error until Reset().
METHOD PRIVATE Move_Timeout_Is_Error
VAR_INST
	rig		: FB_CoverRig;
	nStep	: INT;
	bViol	: BOOL;
END_VAR
TEST('Move_Timeout_Is_Error');
sCurrent := 'Move_Timeout_Is_Error: ';
IF nStep >= 90 THEN
	RETURN;
END_IF
rig.Scan();
CASE nStep OF
0:
	rig.tMoveTimeout := T#300MS;
	rig.fb.Open();
	rig.StepStart();
	nStep := 10;
10:
	IF rig.fb.Error THEN
		Check(rig.StepTime(T#250MS), CONCAT('not before the timeout ', rig.State()));
		Check(rig.OpenOutputs() = '---', CONCAT('the output is off ', rig.State()));
		Check(rig.fb.State = HalfBROT.E_CoverState.Error, CONCAT('state Error after the timeout ', rig.State()));
		rig.fb.Reset();
		nStep := 20;
	ELSIF rig.StepTime(T#2S) THEN
		Check(FALSE, 'no timeout error');
		nStep := 99;
		TEST_FINISHED();
	END_IF
20:
	Check(NOT rig.fb.Error, CONCAT('Reset() clears the timeout error ', rig.State()));
	Check(rig.OpenOutputs() = '---', CONCAT('nothing moves by itself after the reset ', rig.State()));
	nStep := 99;
	TEST_FINISHED();
END_CASE
END_METHOD

// Open() under way, then Close() (#27): the close output waits tReversalDeadTime (300 ms here, 1 s default) after the open output dropped.
METHOD PRIVATE Reversal_Waits_Dead_Time
VAR_INST
	rig		: FB_CoverRig;
	nStep	: INT;
	bViol	: BOOL;
END_VAR
TEST('Reversal_Waits_Dead_Time');
sCurrent := 'Reversal_Waits_Dead_Time: ';
IF nStep >= 90 THEN
	RETURN;
END_IF
rig.Scan();
CASE nStep OF
0:
	rig.tReversalDeadTime := T#300MS;
	rig.fb.Open();
	nStep := 10;
10:
	Check(rig.OpenOutputs() = 'x--', CONCAT('cover 1 opens ', rig.State()));
	rig.SetMid(1);
	rig.fb.Close();
	rig.StepStart();
	nStep := 20;
20:
	Check(rig.OpenOutputs() = '---', CONCAT('the open output is dropped at once ', rig.State()));
	Check(rig.CloseOutputs() = '---', CONCAT('the close output waits for the dead time ', rig.State()));
	nStep := 30;
30:
	bViol := bViol OR (rig.CloseOutputs() <> '---' AND NOT rig.StepTime(T#250MS));
	IF rig.CloseOutputs() <> '---' THEN
		Check(NOT bViol, CONCAT('no close output before the dead time ', rig.State()));
		Check(rig.StepTime(T#250MS) AND NOT rig.StepTime(T#1S), CONCAT('the close output comes after the dead time ', rig.State()));
		Check(rig.CloseOutputs() = 'x--', CONCAT('cover 1 closes ', rig.State()));
		nStep := 99;
		TEST_FINISHED();
	ELSIF rig.StepTime(T#2S) THEN
		Check(FALSE, 'the close output never came');
		nStep := 99;
		TEST_FINISHED();
	END_IF
END_CASE
END_METHOD

END_FUNCTION_BLOCK

// ---- POUs/FB_CoverRig.TcPOU
// FB_CoverControl with limit switches the test sets by hand. The switches are inverted (TRUE = the cover is NOT at the
// switch), see the block: SetClosed(i) puts cover i at its closed switch, SetOpen(i) at its open switch, SetMid(i) between
// them, SetBoth(i) is the limit switch fault (both switches reached). All covers start closed.
// StepStart()/StepTime() measure real time from the start of a step (the block timers run on the system time).
FUNCTION_BLOCK FB_CoverRig
VAR_INPUT
	stIn		: HalfBROT.ST_CoverIn;
	tReversalDeadTime	: TIME := T#1S;
	tMoveTimeout		: TIME := T#60S;
END_VAR
VAR
	fbComm		: FB_NullComm;
	fb			: HalfBROT.FB_CoverControl(comm := fbComm);
	stOut		: HalfBROT.ST_CoverOut;
	tonStep		: TON;
	nScans		: UDINT;
	bInit		: BOOL;
	i			: INT;
END_VAR

METHOD Scan
IF NOT bInit THEN
	bInit := TRUE;
	FOR i := 1 TO 3 DO
		SetClosed(i);
	END_FOR
END_IF
nScans := nScans + 1;
fb(stIn := stIn, tReversalDeadTime := tReversalDeadTime, tMoveTimeout := tMoveTimeout, stOut := stOut);
tonStep(IN := TRUE, PT := T#1H);
END_METHOD

METHOD SetClosed
VAR_INPUT
	nCover	: INT;
END_VAR
stIn.abOpen[nCover] := TRUE;
stIn.abClosed[nCover] := FALSE;
END_METHOD

METHOD SetOpen
VAR_INPUT
	nCover	: INT;
END_VAR
stIn.abOpen[nCover] := FALSE;
stIn.abClosed[nCover] := TRUE;
END_METHOD

METHOD SetMid
VAR_INPUT
	nCover	: INT;
END_VAR
stIn.abOpen[nCover] := TRUE;
stIn.abClosed[nCover] := TRUE;
END_METHOD

METHOD SetBoth
VAR_INPUT
	nCover	: INT;
END_VAR
stIn.abOpen[nCover] := FALSE;
stIn.abClosed[nCover] := FALSE;
END_METHOD

METHOD AllOpen
FOR i := 1 TO 3 DO
	SetOpen(i);
END_FOR
END_METHOD

METHOD AllMid
FOR i := 1 TO 3 DO
	SetMid(i);
END_FOR
END_METHOD

METHOD OpenOutputs : STRING(3)
// the open outputs of cover 1, 2 and 3 as "x" or "-"
OpenOutputs := '';
FOR i := 1 TO 3 DO
	IF stOut.abOpen[i] THEN
		OpenOutputs := CONCAT(OpenOutputs, 'x');
	ELSE
		OpenOutputs := CONCAT(OpenOutputs, '-');
	END_IF
END_FOR
END_METHOD

METHOD CloseOutputs : STRING(3)
// the close outputs of cover 1, 2 and 3 as "x" or "-"
CloseOutputs := '';
FOR i := 1 TO 3 DO
	IF stOut.abClose[i] THEN
		CloseOutputs := CONCAT(CloseOutputs, 'x');
	ELSE
		CloseOutputs := CONCAT(CloseOutputs, '-');
	END_IF
END_FOR
END_METHOD

METHOD State : STRING(60)
State := CONCAT(CONCAT(CONCAT(CONCAT('[open ', OpenOutputs()), ' close '), CloseOutputs()), CONCAT(' err ', BOOL_TO_STRING(fb.bError)));
State := CONCAT(State, ']');
END_METHOD

METHOD StepStart
tonStep(IN := FALSE, PT := T#1H);
END_METHOD

METHOD StepTime : BOOL
VAR_INPUT
	tTime	: TIME;
END_VAR
StepTime := tonStep.ET >= tTime;
END_METHOD

END_FUNCTION_BLOCK

// ---- POUs/FB_PendantControl_Tests.TcPOU
// Characterisation tests of HalfBROT.FB_PendantControl (HalfBROT#32 step 3) through the I/O structs: the selector, the error
// lamp for selector 0 and for blocks that are not connected (#16), the covers (hold-to-run with the key on, the level with the
// key off, #5 cover part) and the hydraulics (start toggle, brake up/down). The focus, derotator, elevation, azimuth and
// telescope selections need their blocks and are only covered for "not connected". They pin what the block does today, they
// are not a specification. Every test owns a rig (FB_PendantRig, the pendant with the cover and hydraulics rigs behind it).
FUNCTION_BLOCK FB_PendantControl_Tests EXTENDS FB_TestBase
VAR
END_VAR

Selector_Decodes_BCD();
Selector_Zero_Lights_Error_Lamp_Only();
Selector_Without_Function_Has_No_Error();
Unset_References_Light_Error_Lamp();
Selector_14_Horn_And_Lamps_Follow_Key();
Cover_Lamps_Show_The_Switches();
Cover_Key_On_Hold_Up_Opens_Release_Stops();
Cover_Key_On_Hold_Down_Closes_Release_Stops();
Cover_Key_On_Up_And_Down_Together_Do_Nothing();
Cover_Run_Stops_When_Selector_Leaves_1_To_3();
Cover_Key_Off_Up_Opens();
Hydraulics_Start_Button_Toggles_Pump();
Hydraulics_Key_Off_Buttons_Do_Nothing();
Hydraulics_Up_Opens_Brake_Down_Closes();

// The four selector inputs are the bits 1, 2, 4 and 8 of Selection.
METHOD PRIVATE Selector_Decodes_BCD
VAR_INST
	rig		: FB_PendantRig;
	nStep	: INT;
	bViol	: BOOL;
END_VAR
TEST('Selector_Decodes_BCD');
sCurrent := 'Selector_Decodes_BCD: ';
IF nStep >= 90 THEN
	RETURN;
END_IF
rig.Scan();
CASE nStep OF
0:
	rig.SetSelector(1);
	rig.StepStart();
	nStep := 10;
10:
	IF rig.nStepScans >= 2 THEN
		Check(rig.fb.Selection = 1, CONCAT('selector 1 ', rig.State()));
		rig.SetSelector(2);
		rig.StepStart();
		nStep := 20;
	END_IF
20:
	IF rig.nStepScans >= 2 THEN
		Check(rig.fb.Selection = 2, CONCAT('selector 2 ', rig.State()));
		rig.SetSelector(4);
		rig.StepStart();
		nStep := 30;
	END_IF
30:
	IF rig.nStepScans >= 2 THEN
		Check(rig.fb.Selection = 4, CONCAT('selector 4 ', rig.State()));
		rig.SetSelector(8);
		rig.StepStart();
		nStep := 40;
	END_IF
40:
	IF rig.nStepScans >= 2 THEN
		Check(rig.fb.Selection = 8, CONCAT('selector 8 ', rig.State()));
		rig.SetSelector(11);
		rig.StepStart();
		nStep := 50;
	END_IF
50:
	IF rig.nStepScans >= 2 THEN
		Check(rig.fb.Selection = 11, CONCAT('selector 11 ', rig.State()));
		rig.SetSelector(15);
		rig.StepStart();
		nStep := 60;
	END_IF
60:
	IF rig.nStepScans >= 2 THEN
		Check(rig.fb.Selection = 15, CONCAT('selector 15 ', rig.State()));
		rig.SetSelector(0);
		rig.StepStart();
		nStep := 70;
	END_IF
70:
	IF rig.nStepScans >= 2 THEN
		Check(rig.fb.Selection = 0, CONCAT('selector 0 ', rig.State()));
		nStep := 99;
		TEST_FINISHED();
	END_IF
END_CASE
END_METHOD

// Selector at 0 (pendant disconnected): only the error lamp, whatever the buttons say; nothing moves (#12).
METHOD PRIVATE Selector_Zero_Lights_Error_Lamp_Only
VAR_INST
	rig		: FB_PendantRig;
	nStep	: INT;
	bViol	: BOOL;
END_VAR
TEST('Selector_Zero_Lights_Error_Lamp_Only');
sCurrent := 'Selector_Zero_Lights_Error_Lamp_Only: ';
IF nStep >= 90 THEN
	RETURN;
END_IF
rig.Scan();
CASE nStep OF
0:
	rig.SetSelector(0); rig.SetKey(TRUE); rig.SetUp(TRUE); rig.SetStart(TRUE);
	rig.StepStart();
	nStep := 10;
10:
	IF rig.nStepScans >= 6 THEN
		Check(rig.Lamps() = '----x', CONCAT('only the error lamp ', rig.State()));
		Check(rig.fb.State = HalfBROT.E_PendantState.Disconnected, CONCAT('state Disconnected ', rig.State()));
		Check(rig.cov.OpenOutputs() = '---' AND rig.cov.CloseOutputs() = '---', CONCAT('no cover moves ', rig.State()));
		Check(NOT rig.hyd.stOut.bOilPumpEnable, CONCAT('no pump ', rig.State()));
		nStep := 99;
		TEST_FINISHED();
	END_IF
END_CASE
END_METHOD

// Selector 4 (Nasmyth), 9 (dome) and 10 (filter wheel) do nothing and light no lamp, also with the key on.
METHOD PRIVATE Selector_Without_Function_Has_No_Error
VAR_INST
	rig		: FB_PendantRig;
	nStep	: INT;
	bViol	: BOOL;
END_VAR
TEST('Selector_Without_Function_Has_No_Error');
sCurrent := 'Selector_Without_Function_Has_No_Error: ';
IF nStep >= 90 THEN
	RETURN;
END_IF
rig.Scan();
CASE nStep OF
0:
	rig.SetKey(TRUE); rig.SetSelector(4);
	rig.StepStart();
	nStep := 10;
10:
	IF rig.nStepScans >= 3 THEN
		Check(rig.Lamps() = '-----', CONCAT('selector 4: no lamp ', rig.State()));
		rig.SetKey(TRUE); rig.SetSelector(9);
		rig.StepStart();
		nStep := 20;
	END_IF
20:
	IF rig.nStepScans >= 3 THEN
		Check(rig.Lamps() = '-----', CONCAT('selector 9: no lamp ', rig.State()));
		rig.SetKey(TRUE); rig.SetSelector(10);
		rig.StepStart();
		nStep := 30;
	END_IF
30:
	IF rig.nStepScans >= 3 THEN
		Check(rig.Lamps() = '-----', CONCAT('selector 10: no lamp ', rig.State()));
		nStep := 99;
		TEST_FINISHED();
	END_IF
END_CASE
END_METHOD

// Selections whose block is not connected (focus, derotator, elevation, azimuth, telescope) light the error lamp and do nothing, with key, start and up pressed: no access to the unset reference (#16).
METHOD PRIVATE Unset_References_Light_Error_Lamp
VAR_INST
	rig		: FB_PendantRig;
	nStep	: INT;
	bViol	: BOOL;
END_VAR
TEST('Unset_References_Light_Error_Lamp');
sCurrent := 'Unset_References_Light_Error_Lamp: ';
IF nStep >= 90 THEN
	RETURN;
END_IF
rig.Scan();
CASE nStep OF
0:
	rig.SetKey(TRUE); rig.SetStart(TRUE); rig.SetUp(TRUE); rig.SetSelector(5);
	rig.StepStart();
	nStep := 10;
10:
	IF rig.nStepScans >= 4 THEN
		Check(rig.Lamps() = '----x', CONCAT('selector 5: block not connected ', rig.State()));
		Check(rig.fb.State = HalfBROT.E_PendantState.ReferencesMissing, CONCAT('state ReferencesMissing ', rig.State()));
		rig.SetKey(TRUE); rig.SetStart(TRUE); rig.SetUp(TRUE); rig.SetSelector(6);
		rig.StepStart();
		nStep := 20;
	END_IF
20:
	IF rig.nStepScans >= 4 THEN
		Check(rig.Lamps() = '----x', CONCAT('selector 6: block not connected ', rig.State()));
		Check(rig.fb.State = HalfBROT.E_PendantState.ReferencesMissing, CONCAT('state ReferencesMissing ', rig.State()));
		rig.SetKey(TRUE); rig.SetStart(TRUE); rig.SetUp(TRUE); rig.SetSelector(7);
		rig.StepStart();
		nStep := 30;
	END_IF
30:
	IF rig.nStepScans >= 4 THEN
		Check(rig.Lamps() = '----x', CONCAT('selector 7: block not connected ', rig.State()));
		Check(rig.fb.State = HalfBROT.E_PendantState.ReferencesMissing, CONCAT('state ReferencesMissing ', rig.State()));
		rig.SetKey(TRUE); rig.SetStart(TRUE); rig.SetUp(TRUE); rig.SetSelector(8);
		rig.StepStart();
		nStep := 40;
	END_IF
40:
	IF rig.nStepScans >= 4 THEN
		Check(rig.Lamps() = '----x', CONCAT('selector 8: block not connected ', rig.State()));
		Check(rig.fb.State = HalfBROT.E_PendantState.ReferencesMissing, CONCAT('state ReferencesMissing ', rig.State()));
		rig.SetKey(TRUE); rig.SetStart(TRUE); rig.SetUp(TRUE); rig.SetSelector(11);
		rig.StepStart();
		nStep := 50;
	END_IF
50:
	IF rig.nStepScans >= 4 THEN
		Check(rig.Lamps() = '----x', CONCAT('selector 11: block not connected ', rig.State()));
		Check(rig.fb.State = HalfBROT.E_PendantState.ReferencesMissing, CONCAT('state ReferencesMissing ', rig.State()));
		rig.SetKey(TRUE); rig.SetStart(TRUE); rig.SetUp(TRUE); rig.SetSelector(12);
		rig.StepStart();
		nStep := 60;
	END_IF
60:
	IF rig.nStepScans >= 4 THEN
		Check(rig.Lamps() = '----x', CONCAT('selector 12: block not connected ', rig.State()));
		Check(rig.fb.State = HalfBROT.E_PendantState.ReferencesMissing, CONCAT('state ReferencesMissing ', rig.State()));
		rig.SetKey(TRUE); rig.SetStart(TRUE); rig.SetUp(TRUE); rig.SetSelector(13);
		rig.StepStart();
		nStep := 70;
	END_IF
70:
	IF rig.nStepScans >= 4 THEN
		Check(rig.Lamps() = '----x', CONCAT('selector 13: block not connected ', rig.State()));
		Check(rig.fb.State = HalfBROT.E_PendantState.ReferencesMissing, CONCAT('state ReferencesMissing ', rig.State()));
		nStep := 99;
		TEST_FINISHED();
	END_IF
END_CASE
END_METHOD

// Selector 14: lamps up, down, left and right and the horn follow the key switch.
METHOD PRIVATE Selector_14_Horn_And_Lamps_Follow_Key
VAR_INST
	rig		: FB_PendantRig;
	nStep	: INT;
	bViol	: BOOL;
END_VAR
TEST('Selector_14_Horn_And_Lamps_Follow_Key');
sCurrent := 'Selector_14_Horn_And_Lamps_Follow_Key: ';
IF nStep >= 90 THEN
	RETURN;
END_IF
rig.Scan();
CASE nStep OF
0:
	rig.SetSelector(14);
	rig.StepStart();
	nStep := 10;
10:
	IF rig.nStepScans >= 3 THEN
		Check(rig.Lamps() = '-----', CONCAT('key off: no lamp ', rig.State()));
		Check(rig.fb.State = HalfBROT.E_PendantState.Automatic, CONCAT('key off: state Automatic ', rig.State()));
		Check(NOT rig.fb.horn, CONCAT('key off: no horn ', rig.State()));
		rig.SetKey(TRUE);
		rig.StepStart();
		nStep := 20;
	END_IF
20:
	IF rig.nStepScans >= 3 THEN
		Check(rig.Lamps() = 'xxxx-', CONCAT('key on: four lamps, no error lamp ', rig.State()));
		Check(rig.fb.State = HalfBROT.E_PendantState.Manual, CONCAT('key on: state Manual ', rig.State()));
		Check(rig.fb.horn, CONCAT('key on: horn ', rig.State()));
		rig.SetKey(FALSE);
		rig.StepStart();
		nStep := 30;
	END_IF
30:
	IF rig.nStepScans >= 3 THEN
		Check(rig.Lamps() = '-----', CONCAT('key off again: no lamp ', rig.State()));
		Check(NOT rig.fb.horn, CONCAT('key off again: no horn ', rig.State()));
		nStep := 99;
		TEST_FINISHED();
	END_IF
END_CASE
END_METHOD

// Selector 1: up is lit while the cover is not at its open switch, down while it is not at its closed switch; with the key on the error lamp shows a limit switch fault.
METHOD PRIVATE Cover_Lamps_Show_The_Switches
VAR_INST
	rig		: FB_PendantRig;
	nStep	: INT;
	bViol	: BOOL;
END_VAR
TEST('Cover_Lamps_Show_The_Switches');
sCurrent := 'Cover_Lamps_Show_The_Switches: ';
IF nStep >= 90 THEN
	RETURN;
END_IF
rig.Scan();
CASE nStep OF
0:
	rig.SetSelector(1);
	rig.StepStart();
	nStep := 10;
10:
	IF rig.nStepScans >= 5 THEN
		Check(rig.Lamps() = 'x----', CONCAT('closed: up lit, down dark ', rig.State()));
		rig.cov.AllOpen();
		rig.StepStart();
		nStep := 20;
	END_IF
20:
	IF rig.nStepScans >= 5 THEN
		Check(rig.Lamps() = '-x---', CONCAT('open: up dark, down lit ', rig.State()));
		rig.cov.SetBoth(1); rig.SetKey(TRUE);
		rig.StepStart();
		nStep := 30;
	END_IF
30:
	IF rig.nStepScans >= 5 THEN
		Check(rig.Lamps() = '----x', CONCAT('both switches reached: error lamp ', rig.State()));
		rig.cov.SetMid(1);
		rig.StepStart();
		nStep := 40;
	END_IF
40:
	IF rig.nStepScans >= 5 THEN
		Check(rig.Lamps() = 'xx---', CONCAT('between the switches: up and down lit, no error ', rig.State()));
		nStep := 99;
		TEST_FINISHED();
	END_IF
END_CASE
END_METHOD

// Key on, selector 1: up held opens cover 1 (the block does the order); releasing the button stops the run.
METHOD PRIVATE Cover_Key_On_Hold_Up_Opens_Release_Stops
VAR_INST
	rig		: FB_PendantRig;
	nStep	: INT;
	bViol	: BOOL;
END_VAR
TEST('Cover_Key_On_Hold_Up_Opens_Release_Stops');
sCurrent := 'Cover_Key_On_Hold_Up_Opens_Release_Stops: ';
IF nStep >= 90 THEN
	RETURN;
END_IF
rig.Scan();
CASE nStep OF
0:
	rig.SetSelector(1); rig.SetKey(TRUE);
	rig.StepStart();
	nStep := 10;
10:
	IF rig.nStepScans >= 4 THEN
		Check(rig.cov.OpenOutputs() = '---' AND rig.cov.CloseOutputs() = '---', CONCAT('nothing moves without a button ', rig.State()));
		rig.SetUp(TRUE);
		rig.StepStart();
		nStep := 20;
	END_IF
20:
	IF rig.nStepScans >= 25 THEN
		Check(rig.cov.OpenOutputs() = 'x--' AND rig.cov.CloseOutputs() = '---', CONCAT('up held: cover 1 opens ', rig.State()));
		rig.SetUp(FALSE);
		rig.StepStart();
		nStep := 30;
	END_IF
30:
	IF rig.nStepScans >= 25 THEN
		Check(rig.cov.OpenOutputs() = '---' AND rig.cov.CloseOutputs() = '---', CONCAT('the release stops the run ', rig.State()));
		nStep := 99;
		TEST_FINISHED();
	END_IF
END_CASE
END_METHOD

// Key on, selector 1, all covers open: down held closes cover 2 first; releasing the button stops the run.
METHOD PRIVATE Cover_Key_On_Hold_Down_Closes_Release_Stops
VAR_INST
	rig		: FB_PendantRig;
	nStep	: INT;
	bViol	: BOOL;
END_VAR
TEST('Cover_Key_On_Hold_Down_Closes_Release_Stops');
sCurrent := 'Cover_Key_On_Hold_Down_Closes_Release_Stops: ';
IF nStep >= 90 THEN
	RETURN;
END_IF
rig.Scan();
CASE nStep OF
0:
	rig.cov.AllOpen(); rig.SetSelector(1); rig.SetKey(TRUE);
	rig.StepStart();
	nStep := 10;
10:
	IF rig.nStepScans >= 5 THEN
		Check(rig.cov.OpenOutputs() = '---' AND rig.cov.CloseOutputs() = '---', CONCAT('nothing moves without a button ', rig.State()));
		rig.SetDown(TRUE);
		rig.StepStart();
		nStep := 20;
	END_IF
20:
	IF rig.nStepScans >= 25 THEN
		Check(rig.cov.CloseOutputs() = '-x-' AND rig.cov.OpenOutputs() = '---', CONCAT('down held: cover 2 closes first ', rig.State()));
		rig.SetDown(FALSE);
		rig.StepStart();
		nStep := 30;
	END_IF
30:
	IF rig.nStepScans >= 5 THEN
		Check(rig.cov.OpenOutputs() = '---' AND rig.cov.CloseOutputs() = '---', CONCAT('the release stops the run ', rig.State()));
		nStep := 99;
		TEST_FINISHED();
	END_IF
END_CASE
END_METHOD

// Key on, selector 1: up and down pressed together start nothing.
METHOD PRIVATE Cover_Key_On_Up_And_Down_Together_Do_Nothing
VAR_INST
	rig		: FB_PendantRig;
	nStep	: INT;
	bViol	: BOOL;
END_VAR
TEST('Cover_Key_On_Up_And_Down_Together_Do_Nothing');
sCurrent := 'Cover_Key_On_Up_And_Down_Together_Do_Nothing: ';
IF nStep >= 90 THEN
	RETURN;
END_IF
rig.Scan();
CASE nStep OF
0:
	rig.SetSelector(1); rig.SetKey(TRUE); rig.SetUp(TRUE); rig.SetDown(TRUE);
	rig.StepStart();
	nStep := 10;
10:
	IF rig.nStepScans >= 12 THEN
		Check(rig.cov.OpenOutputs() = '---' AND rig.cov.CloseOutputs() = '---', CONCAT('up and down together ', rig.State()));
		nStep := 99;
		TEST_FINISHED();
	END_IF
END_CASE
END_METHOD

// A run started by the pendant stops when the selector leaves 1 to 3 although the button is still held.
METHOD PRIVATE Cover_Run_Stops_When_Selector_Leaves_1_To_3
VAR_INST
	rig		: FB_PendantRig;
	nStep	: INT;
	bViol	: BOOL;
END_VAR
TEST('Cover_Run_Stops_When_Selector_Leaves_1_To_3');
sCurrent := 'Cover_Run_Stops_When_Selector_Leaves_1_To_3: ';
IF nStep >= 90 THEN
	RETURN;
END_IF
rig.Scan();
CASE nStep OF
0:
	rig.SetSelector(1); rig.SetKey(TRUE); rig.SetUp(TRUE);
	rig.StepStart();
	nStep := 10;
10:
	IF rig.nStepScans >= 6 THEN
		Check(rig.cov.OpenOutputs() = 'x--', CONCAT('cover 1 opens ', rig.State()));
		rig.SetSelector(4);
		rig.StepStart();
		nStep := 20;
	END_IF
20:
	IF rig.nStepScans >= 4 THEN
		Check(rig.cov.OpenOutputs() = '---' AND rig.cov.CloseOutputs() = '---', CONCAT('the run stops with the selector ', rig.State()));
		nStep := 99;
		TEST_FINISHED();
	END_IF
END_CASE
END_METHOD

// Key off (automatic), selector 1: up opens cover 1 (the level, no hold-to-run).
METHOD PRIVATE Cover_Key_Off_Up_Opens
VAR_INST
	rig		: FB_PendantRig;
	nStep	: INT;
	bViol	: BOOL;
END_VAR
TEST('Cover_Key_Off_Up_Opens');
sCurrent := 'Cover_Key_Off_Up_Opens: ';
IF nStep >= 90 THEN
	RETURN;
END_IF
rig.Scan();
CASE nStep OF
0:
	rig.SetSelector(1); rig.SetUp(TRUE);
	rig.StepStart();
	nStep := 10;
10:
	IF rig.nStepScans >= 6 THEN
		Check(rig.cov.OpenOutputs() = 'x--' AND rig.cov.CloseOutputs() = '---', CONCAT('up: cover 1 opens ', rig.State()));
		nStep := 99;
		TEST_FINISHED();
	END_IF
END_CASE
END_METHOD

// Key on, selector 15: each press of start (the edge, not the level) toggles the hydraulics enable; the lamps show pump and pressure.
METHOD PRIVATE Hydraulics_Start_Button_Toggles_Pump
VAR_INST
	rig		: FB_PendantRig;
	nStep	: INT;
	bViol	: BOOL;
END_VAR
TEST('Hydraulics_Start_Button_Toggles_Pump');
sCurrent := 'Hydraulics_Start_Button_Toggles_Pump: ';
IF nStep >= 90 THEN
	RETURN;
END_IF
rig.Scan();
CASE nStep OF
0:
	rig.SetSelector(15); rig.SetKey(TRUE);
	rig.StepStart();
	nStep := 10;
10:
	IF rig.nStepScans >= 4 THEN
		Check(NOT rig.hyd.stOut.bOilPumpEnable, CONCAT('the pump is off ', rig.State()));
		rig.SetStart(TRUE);
		rig.StepStart();
		nStep := 20;
	END_IF
20:
	IF rig.nStepScans >= 15 THEN
		Check(rig.hyd.stOut.bOilPumpEnable AND rig.hyd.fb.Enable, CONCAT('the pump is enabled ', rig.State()));
		Check(rig.hyd.fb.PumpRunning AND rig.hyd.fb.OilPressureOK, CONCAT('pump running with pressure ', rig.State()));
		Check(rig.stOut.bLampLeft AND rig.stOut.bLampUp AND NOT rig.stOut.bLampDown, CONCAT('lamps: pump running, pressure, brake closed ', rig.State()));
		rig.SetStart(FALSE);
		rig.StepStart();
		nStep := 30;
	END_IF
30:
	IF rig.nStepScans >= 8 THEN
		Check(rig.hyd.stOut.bOilPumpEnable AND rig.hyd.fb.Enable, CONCAT('the pump is still enabled after the button was held and released ', rig.State()));
		rig.SetStart(TRUE);
		rig.StepStart();
		nStep := 40;
	END_IF
40:
	IF rig.nStepScans >= 8 THEN
		Check(NOT rig.hyd.stOut.bOilPumpEnable AND NOT rig.hyd.fb.Enable, CONCAT('the second press stops the pump ', rig.State()));
		rig.SetStart(FALSE);
		rig.StepStart();
		nStep := 50;
	END_IF
50:
	IF rig.nStepScans >= 6 THEN
		Check(NOT rig.stOut.bLampLeft AND NOT rig.stOut.bLampUp, CONCAT('lamps: pump stopped ', rig.State()));
		nStep := 99;
		TEST_FINISHED();
	END_IF
END_CASE
END_METHOD

// Key off, selector 15: start and up change nothing (the buttons work with the key on only).
METHOD PRIVATE Hydraulics_Key_Off_Buttons_Do_Nothing
VAR_INST
	rig		: FB_PendantRig;
	nStep	: INT;
	bViol	: BOOL;
END_VAR
TEST('Hydraulics_Key_Off_Buttons_Do_Nothing');
sCurrent := 'Hydraulics_Key_Off_Buttons_Do_Nothing: ';
IF nStep >= 90 THEN
	RETURN;
END_IF
rig.Scan();
CASE nStep OF
0:
	rig.SetSelector(15); rig.SetStart(TRUE); rig.SetUp(TRUE);
	rig.StepStart();
	nStep := 10;
10:
	IF rig.nStepScans >= 15 THEN
		Check(NOT rig.hyd.stOut.bOilPumpEnable AND NOT rig.hyd.fb.Enable, CONCAT('no pump ', rig.State()));
		Check(NOT rig.stOut.bLampLeft AND NOT rig.stOut.bLampUp AND NOT rig.stOut.bLampDown, CONCAT('no lamp ', rig.State()));
		nStep := 99;
		TEST_FINISHED();
	END_IF
END_CASE
END_METHOD

// Key on, selector 15, pump running: up held opens the brake (pressure delay 3 s), down closes it; the lamps follow.
METHOD PRIVATE Hydraulics_Up_Opens_Brake_Down_Closes
VAR_INST
	rig		: FB_PendantRig;
	nStep	: INT;
	bViol	: BOOL;
END_VAR
TEST('Hydraulics_Up_Opens_Brake_Down_Closes');
sCurrent := 'Hydraulics_Up_Opens_Brake_Down_Closes: ';
IF nStep >= 90 THEN
	RETURN;
END_IF
rig.Scan();
CASE nStep OF
0:
	rig.SetSelector(15);
	rig.SetKey(TRUE);
	rig.SetClearing(TRUE);
	rig.SetStart(TRUE);
	rig.StepStart();
	nStep := 10;
10:
	IF rig.nStepScans >= 3 THEN
		rig.SetStart(FALSE);
		rig.StepStart();
		nStep := 20;
	END_IF
20:
	IF rig.hyd.fb.OilPressureOK THEN
		rig.SetUp(TRUE);
		rig.StepStart();
		nStep := 30;
	ELSIF rig.StepTime(T#2S) THEN
		Check(FALSE, 'the pump did not come up');
		nStep := 99;
		TEST_FINISHED();
	END_IF
30:
	IF rig.hyd.fb.BrakeOpen THEN
		rig.StepStart();
		nStep := 35;
	ELSIF rig.StepTime(T#8S) THEN
		Check(FALSE, 'up held did not open the brake');
		nStep := 99;
		TEST_FINISHED();
	END_IF
35:
	IF rig.nStepScans >= 3 THEN
		Check(rig.stOut.bLampDown AND NOT rig.stOut.bLampUp, CONCAT('lamps: pressure, brake open ', rig.State()));
		rig.SetUp(FALSE);
		rig.SetDown(TRUE);
		rig.StepStart();
		nStep := 40;
	END_IF
40:
	IF NOT rig.hyd.fb.BrakeOpen THEN
		Check(NOT rig.hyd.stOut.bBrakeAzEl, CONCAT('the brake output is off ', rig.State()));
		rig.StepStart();
		nStep := 45;
	ELSIF rig.StepTime(T#1S) THEN
		Check(FALSE, 'down held did not close the brake');
		nStep := 99;
		TEST_FINISHED();
	END_IF
45:
	IF rig.nStepScans >= 3 THEN
		Check(rig.stOut.bLampUp AND NOT rig.stOut.bLampDown, CONCAT('lamps: pressure, brake closed ', rig.State()));
		nStep := 99;
		TEST_FINISHED();
	END_IF
END_CASE
END_METHOD

END_FUNCTION_BLOCK

// ---- POUs/FB_PendantRig.TcPOU
// FB_PendantControl with the cover block and the hydraulics block behind it, each in its rig (FB_CoverRig, FB_HydraulicsRig).
// The other blocks the pendant can reference (focus, elevation, azimuth, derotator, telescope) are not connected: the pendant
// must light the error lamp and do nothing for those selections (#16). The test sets the pendant inputs through SetKey(),
// SetSelector(), SetUp() ... and reads the lamps through Lamps() ("x" = lit, order up, down, left, right, error).
// The pendant runs before the blocks in every scan, like in MAIN. StepStart()/nStepScans count the scans from the start of a step.
FUNCTION_BLOCK FB_PendantRig
VAR_INPUT
	stIn		: HalfBROT.ST_PendantIn;
END_VAR
VAR
	fbComm		: FB_NullComm;
	fb			: HalfBROT.FB_PendantControl(comm := fbComm);
	stOut		: HalfBROT.ST_PendantOut;
	cov			: FB_CoverRig;
	hyd			: FB_HydraulicsRig;
	tonStep		: TON;
	nScans		: UDINT;
	nStepScans	: UDINT;
END_VAR

METHOD Scan
nScans := nScans + 1;
nStepScans := nStepScans + 1;
fb(stIn := stIn, fbCovers := cov.fb, fbBrake := hyd.fb, fbHydraulics := hyd.fb, stOut := stOut);
cov.Scan();
hyd.Scan();
tonStep(IN := TRUE, PT := T#1H);
END_METHOD

METHOD SetKey
VAR_INPUT
	bOn	: BOOL;
END_VAR
stIn.bKeySwitch := bOn;
END_METHOD

METHOD SetUp
VAR_INPUT
	bOn	: BOOL;
END_VAR
stIn.bDirectionUp := bOn;
END_METHOD

METHOD SetDown
VAR_INPUT
	bOn	: BOOL;
END_VAR
stIn.bDirectionDown := bOn;
END_METHOD

METHOD SetLeft
VAR_INPUT
	bOn	: BOOL;
END_VAR
stIn.bDirectionLeft := bOn;
END_METHOD

METHOD SetRight
VAR_INPUT
	bOn	: BOOL;
END_VAR
stIn.bDirectionRight := bOn;
END_METHOD

METHOD SetStart
VAR_INPUT
	bOn	: BOOL;
END_VAR
stIn.bStartSwitch := bOn;
END_METHOD

METHOD SetReset
VAR_INPUT
	bOn	: BOOL;
END_VAR
stIn.bResetSwitch := bOn;
END_METHOD

METHOD SetSelector
VAR_INPUT
	nSelector	: INT;
END_VAR
stIn.bBCD0 := (nSelector AND 1) <> 0;
stIn.bBCD2 := (nSelector AND 2) <> 0;
stIn.bBCD4 := (nSelector AND 4) <> 0;
stIn.bBCD8 := (nSelector AND 8) <> 0;
END_METHOD

METHOD SetClearing
VAR_INPUT
	bOn	: BOOL;
END_VAR
hyd.bClearing := bOn;
END_METHOD

METHOD Lamps : STRING(5)
Lamps := '';
IF stOut.bLampUp THEN
	Lamps := CONCAT(Lamps, 'x');
ELSE
	Lamps := CONCAT(Lamps, '-');
END_IF
IF stOut.bLampDown THEN
	Lamps := CONCAT(Lamps, 'x');
ELSE
	Lamps := CONCAT(Lamps, '-');
END_IF
IF stOut.bLampLeft THEN
	Lamps := CONCAT(Lamps, 'x');
ELSE
	Lamps := CONCAT(Lamps, '-');
END_IF
IF stOut.bLampRight THEN
	Lamps := CONCAT(Lamps, 'x');
ELSE
	Lamps := CONCAT(Lamps, '-');
END_IF
IF stOut.bLampError THEN
	Lamps := CONCAT(Lamps, 'x');
ELSE
	Lamps := CONCAT(Lamps, '-');
END_IF
END_METHOD

METHOD State : STRING(100)
State := CONCAT('[sel ', UINT_TO_STRING(fb.Selection));
State := CONCAT(State, CONCAT(' lamps ', Lamps()));
State := CONCAT(State, CONCAT(' open ', cov.OpenOutputs()));
State := CONCAT(State, CONCAT(' close ', cov.CloseOutputs()));
State := CONCAT(State, CONCAT(' pump ', BOOL_TO_STRING(hyd.stOut.bOilPumpEnable)));
State := CONCAT(State, ']');
END_METHOD

METHOD StepStart
tonStep(IN := FALSE, PT := T#1H);
nStepScans := 0;
END_METHOD

METHOD StepTime : BOOL
VAR_INPUT
	tTime	: TIME;
END_VAR
StepTime := tonStep.ET >= tTime;
END_METHOD

END_FUNCTION_BLOCK

// ---- POUs/FB_FocusUnlock_Tests.TcPOU
// Unlock sequence of the focus (HalfBROT.FB_FocusUnlock, wired into FB_FocusControl): the drive is powered while the lock
// is closed, the lock opens only after the power status, no move before ptFocusDelay after the unlock, a power timeout
// keeps the lock closed (until Reset), an error and a dropped request close the lock and drop the drive in one cycle.
// Every test owns a rig (FB_FocusUnlockRig: drive model + the real FB_MoveFollower) and runs over several PLC cycles
// in real time (power up 200 ms, settle 50 ms, focus delay 300 ms unless the test sets other times).
FUNCTION_BLOCK FB_FocusUnlock_Tests EXTENDS FB_TestBase
VAR
END_VAR

Lock_Opens_Only_After_Power_Status();
No_Move_Before_Focus_Delay();
Power_Timeout_Keeps_Lock_Closed();
Power_Lost_Closes_Lock();
Error_Closes_Lock_And_Drops_Drive_In_One_Cycle();
Request_Drop_Locks_In_One_Cycle();

// The request enables the drive at once with the lock closed; the lock opens only after the power status (200 ms) and
// the settle time (50 ms), and bUnlocked (moves allowed) is still FALSE then.
METHOD PRIVATE Lock_Opens_Only_After_Power_Status
VAR_INST
	rig		: FB_FocusUnlockRig;
	nStep	: INT;
	bViol	: BOOL;
END_VAR
TEST('Lock_Opens_Only_After_Power_Status');
sCurrent := 'Lock_Opens_Only_After_Power_Status: ';
IF nStep >= 90 THEN
	RETURN;
END_IF
CASE nStep OF
0:
	rig.bRequest := TRUE;
	rig.StepStart();
	rig.Scan();
	Check(rig.fb.bDriveEnable, CONCAT('the drive is enabled with the request ', rig.State()));
	Check(NOT rig.fb.bUnlock, CONCAT('the lock stays closed until the drive reports power ', rig.State()));
	nStep := 10;
10:
	rig.Scan();
	bViol := bViol OR (rig.fb.bUnlock AND NOT rig.bPowered) OR NOT rig.fb.bDriveEnable;
	IF rig.fb.bUnlock THEN
		Check(NOT bViol, CONCAT('no unlock without power status, the drive stays enabled ', rig.State()));
		Check(rig.StepTime(T#240MS), CONCAT('the lock opens after power up and settle time ', rig.State()));
		Check(NOT rig.fb.bUnlocked, CONCAT('no move allowed in the cycle the lock opens ', rig.State()));
		nStep := 99;
		TEST_FINISHED();
	ELSIF rig.StepTime(T#2S) THEN
		Check(FALSE, CONCAT('the lock never opened ', rig.State()));
		nStep := 99;
		TEST_FINISHED();
	END_IF
END_CASE
END_METHOD

// Automatic positioning with the focus off its target: the follower starts the move only when the lock has been open for
// tFocusDelay (300 ms), never while the lock is closed or still releasing.
METHOD PRIVATE No_Move_Before_Focus_Delay
VAR_INST
	rig		: FB_FocusUnlockRig;
	nStep	: INT;
END_VAR
TEST('No_Move_Before_Focus_Delay');
sCurrent := 'No_Move_Before_Focus_Delay: ';
IF nStep >= 90 THEN
	RETURN;
END_IF
CASE nStep OF
0:
	rig.bFollow := TRUE;
	rig.bRequest := TRUE;
	rig.StepStart();
	rig.Scan();
	nStep := 10;
10:
	rig.Scan();
	IF rig.nStarts > 0 THEN
		Check(NOT rig.bStartBeforeUnlocked, CONCAT('no move before bUnlocked ', rig.State()));
		Check(rig.tUnlockAt < T#1H, CONCAT('the lock is open ', rig.State()));
		Check(rig.tFirstStart >= rig.tUnlockAt + T#280MS, CONCAT('the move starts ptFocusDelay after the unlock ', rig.State()));
		Check(rig.tFirstStart <= rig.tUnlockAt + T#500MS, CONCAT('and not much later ', rig.State()));
		nStep := 99;
		TEST_FINISHED();
	ELSIF rig.StepTime(T#2S) THEN
		Check(FALSE, CONCAT('the move never started ', rig.State()));
		nStep := 99;
		TEST_FINISHED();
	END_IF
END_CASE
END_METHOD

// The drive never reports power: after tPowerTimeout (400 ms here) bPowerTimeout, the drive is dropped and the lock never
// opened. It stays so until Reset; after the reset the sequence runs again and unlocks once the drive powers.
METHOD PRIVATE Power_Timeout_Keeps_Lock_Closed
VAR_INST
	rig		: FB_FocusUnlockRig;
	nStep	: INT;
	bViol	: BOOL;
END_VAR
TEST('Power_Timeout_Keeps_Lock_Closed');
sCurrent := 'Power_Timeout_Keeps_Lock_Closed: ';
IF nStep >= 90 THEN
	RETURN;
END_IF
CASE nStep OF
0:
	rig.bDrivePowers := FALSE;
	rig.tPowerTimeout := T#400MS;
	rig.bFollow := TRUE;
	rig.bRequest := TRUE;
	rig.StepStart();
	rig.Scan();
	nStep := 10;
10:
	rig.Scan();
	bViol := bViol OR rig.fb.bUnlock OR rig.nStarts > 0;
	IF rig.StepTime(T#800MS) THEN
		Check(NOT bViol, CONCAT('the lock never opened, no move ', rig.State()));
		Check(rig.fb.bPowerTimeout, CONCAT('power timeout ', rig.State()));
		Check(rig.tTimeoutAt >= T#380MS AND rig.tTimeoutAt <= T#600MS, CONCAT('after tPowerTimeout ', rig.State()));
		Check(NOT rig.fb.bDriveEnable, CONCAT('the drive is dropped ', rig.State()));
		rig.bReset := TRUE;
		nStep := 20;
	END_IF
20:
	rig.Scan();
	rig.bReset := FALSE;
	Check(NOT rig.fb.bPowerTimeout, CONCAT('Reset clears the timeout ', rig.State()));
	Check(rig.fb.bDriveEnable AND NOT rig.fb.bUnlock, CONCAT('the drive is enabled again, lock closed ', rig.State()));
	rig.bDrivePowers := TRUE;
	rig.StepStart();
	nStep := 30;
30:
	rig.Scan();
	IF rig.fb.bUnlock THEN
		Check(rig.bPowered AND NOT rig.fb.bPowerTimeout, CONCAT('unlocked with power after the reset ', rig.State()));
		nStep := 99;
		TEST_FINISHED();
	ELSIF rig.StepTime(T#2S) THEN
		Check(FALSE, CONCAT('no unlock after the reset ', rig.State()));
		nStep := 99;
		TEST_FINISHED();
	END_IF
END_CASE
END_METHOD

// Unlocked, then the drive loses its power status without an axis error: the lock closes in the next cycle, no move is
// allowed, and it is a power timeout after tPowerTimeout (400 ms here).
METHOD PRIVATE Power_Lost_Closes_Lock
VAR_INST
	rig		: FB_FocusUnlockRig;
	nStep	: INT;
	bViol	: BOOL;
END_VAR
TEST('Power_Lost_Closes_Lock');
sCurrent := 'Power_Lost_Closes_Lock: ';
IF nStep >= 90 THEN
	RETURN;
END_IF
CASE nStep OF
0:
	rig.tPowerTimeout := T#400MS;
	rig.bRequest := TRUE;
	rig.StepStart();
	rig.Scan();
	nStep := 10;
10:
	rig.Scan();
	IF rig.fb.bUnlocked THEN
		rig.bDrivePowers := FALSE;	// takes effect in the "fbAxis call" of the next Scan
		nStep := 20;
	ELSIF rig.StepTime(T#2S) THEN
		Check(FALSE, CONCAT('never unlocked ', rig.State()));
		nStep := 99;
		TEST_FINISHED();
	END_IF
20:
	rig.Scan();		// power status drops in this fbAxis call
	rig.Scan();		// the unlock sequence sees it
	Check(NOT rig.fb.bUnlock AND NOT rig.fb.bUnlocked, CONCAT('the lock closes when the power status is lost ', rig.State()));
	rig.StepStart();
	nStep := 30;
30:
	rig.Scan();
	bViol := bViol OR rig.fb.bUnlock;
	IF rig.StepTime(T#700MS) THEN
		Check(NOT bViol, CONCAT('the lock stays closed ', rig.State()));
		Check(rig.fb.bPowerTimeout AND NOT rig.fb.bDriveEnable, CONCAT('power timeout, drive dropped ', rig.State()));
		nStep := 99;
		TEST_FINISHED();
	END_IF
END_CASE
END_METHOD

// Unlocked and ready to move, then an axis error: the first call that sees bError closes the lock and drops the drive
// (and bUnlocked). After the error is gone the sequence starts again with the lock closed.
METHOD PRIVATE Error_Closes_Lock_And_Drops_Drive_In_One_Cycle
VAR_INST
	rig		: FB_FocusUnlockRig;
	nStep	: INT;
END_VAR
TEST('Error_Closes_Lock_And_Drops_Drive_In_One_Cycle');
sCurrent := 'Error_Closes_Lock_And_Drops_Drive_In_One_Cycle: ';
IF nStep >= 90 THEN
	RETURN;
END_IF
CASE nStep OF
0:
	rig.bRequest := TRUE;
	rig.StepStart();
	rig.Scan();
	nStep := 10;
10:
	rig.Scan();
	IF rig.fb.bUnlocked THEN
		rig.bError := TRUE;
		rig.Scan();
		Check(NOT rig.fb.bUnlock, CONCAT('the lock closes in the error cycle ', rig.State()));
		Check(NOT rig.fb.bDriveEnable, CONCAT('the drive drops in the error cycle ', rig.State()));
		Check(NOT rig.fb.bUnlocked, CONCAT('no move allowed ', rig.State()));
		Check(NOT rig.fb.bPowerTimeout, CONCAT('an axis error is no power timeout ', rig.State()));
		rig.bError := FALSE;
		rig.Scan();
		Check(rig.fb.bDriveEnable AND NOT rig.fb.bUnlock, CONCAT('after the error: drive first, lock closed ', rig.State()));
		nStep := 99;
		TEST_FINISHED();
	ELSIF rig.StepTime(T#2S) THEN
		Check(FALSE, CONCAT('never unlocked ', rig.State()));
		nStep := 99;
		TEST_FINISHED();
	END_IF
END_CASE
END_METHOD

// Locking is unchanged: when the request drops (FB_FocusDriveEnable after ptBrakeDelay, or bManualUnlock off) the lock
// closes and the drive drops in the same cycle.
METHOD PRIVATE Request_Drop_Locks_In_One_Cycle
VAR_INST
	rig		: FB_FocusUnlockRig;
	nStep	: INT;
END_VAR
TEST('Request_Drop_Locks_In_One_Cycle');
sCurrent := 'Request_Drop_Locks_In_One_Cycle: ';
IF nStep >= 90 THEN
	RETURN;
END_IF
CASE nStep OF
0:
	rig.bRequest := TRUE;
	rig.StepStart();
	rig.Scan();
	nStep := 10;
10:
	rig.Scan();
	IF rig.fb.bUnlocked THEN
		rig.bRequest := FALSE;
		rig.Scan();
		Check(NOT rig.fb.bUnlock AND NOT rig.fb.bDriveEnable AND NOT rig.fb.bUnlocked,
			CONCAT('lock closed and drive off together ', rig.State()));
		nStep := 99;
		TEST_FINISHED();
	ELSIF rig.StepTime(T#2S) THEN
		Check(FALSE, CONCAT('never unlocked ', rig.State()));
		nStep := 99;
		TEST_FINISHED();
	END_IF
END_CASE
END_METHOD

END_FUNCTION_BLOCK

// ---- POUs/FB_FocusUnlockRig.TcPOU
// HalfBROT.FB_FocusUnlock in the order of FB_FocusControl, with a drive model and the real BROTLib.FB_MoveFollower behind
// it: Scan() is one PLC cycle (unlock sequence, follower, then the "fbAxis call": the power status comes tPowerUp after
// the enable, never with bDrivePowers FALSE, and drops with the enable). The follower gets bReady as in FB_FocusControl
// (fbAxis.Ready AND bFocusUnlocked AND bEnable) and is active with bFollow; the axis does not move, a start is counted.
// tUnlockAt / tFirstStart: the step time of the first cycle with the lock open / with a move started (T#1H = not yet).
// StepStart()/StepTime() measure real time from the start of a step (the block timers run on the system time).
FUNCTION_BLOCK FB_FocusUnlockRig
VAR_INPUT
	bRequest		: BOOL;		// bManualUnlock OR bEnable
	bError			: BOOL;
	bReset			: BOOL;
	bDrivePowers	: BOOL := TRUE;		// FALSE: the power status never comes
	bFollow			: BOOL;		// automatic positioning (follower active)
	fTarget			: LREAL := 10.0;
	fActual			: LREAL := 8.0;
	tPowerUp		: TIME := T#200MS;	// enable -> power status of the drive model
	tPowerSettle	: TIME := T#50MS;
	tPowerTimeout	: TIME := T#2S;
	tFocusDelay		: TIME := T#300MS;
END_VAR
VAR_OUTPUT
	bPowered		: BOOL;		// fbAxis.Ready of the last "fbAxis call"
	nStarts			: INT;		// cycles with bStartMove
	bStartBeforeUnlocked	: BOOL;	// a move started while bUnlocked was FALSE
	tUnlockAt		: TIME := T#1H;
	tFirstStart		: TIME := T#1H;
	tTimeoutAt		: TIME := T#1H;	// first cycle with bPowerTimeout
END_VAR
VAR
	fb				: HalfBROT.FB_FocusUnlock;
	fbFollower		: BROTLib.FB_MoveFollower;
	tonPowerUp		: TON;
	tonStep			: TON;
END_VAR

METHOD Scan
fb(
	bRequest		:= bRequest,
	bError			:= bError,
	bPowered		:= bPowered,
	bReset			:= bReset,
	tPowerSettle	:= tPowerSettle,
	tPowerTimeout	:= tPowerTimeout,
	tFocusDelay		:= tFocusDelay);
IF fb.bUnlock AND tUnlockAt = T#1H THEN
	tUnlockAt := tonStep.ET;
END_IF
IF fb.bPowerTimeout AND tTimeoutAt = T#1H THEN
	tTimeoutAt := tonStep.ET;
END_IF

fbFollower(
	fTarget		:= fTarget,
	fActual		:= fActual,
	fTolerance	:= 0.005,
	bActive		:= bFollow,
	bReady		:= bPowered AND fb.bUnlocked AND bRequest,
	bMoveDone	:= FALSE,
	bAborted	:= FALSE,
	bError		:= bError,
	bStopDone	:= FALSE);
IF fbFollower.bStartMove THEN
	nStarts := nStarts + 1;
	bStartBeforeUnlocked := bStartBeforeUnlocked OR NOT fb.bUnlocked OR NOT fb.bUnlock;
	IF tFirstStart = T#1H THEN
		tFirstStart := tonStep.ET;
	END_IF
END_IF

// the "fbAxis call": MC_Power gets fb.bDriveEnable
tonPowerUp(IN := fb.bDriveEnable AND bDrivePowers, PT := tPowerUp);
bPowered := tonPowerUp.Q;

tonStep(IN := TRUE, PT := T#1H);
END_METHOD

METHOD StepStart
tonStep(IN := FALSE, PT := T#1H);
tUnlockAt := T#1H;
tFirstStart := T#1H;
tTimeoutAt := T#1H;
END_METHOD

METHOD StepTime : BOOL
VAR_INPUT
	tTime	: TIME;
END_VAR
StepTime := tonStep.ET >= tTime;
END_METHOD

// 'enable=1 powered=0 unlock=0 unlocked=0 timeout=0 starts=0' for the failure texts
METHOD State : STRING(255)
State := CONCAT('enable=', BOOL_TO_STRING(fb.bDriveEnable));
State := CONCAT(State, CONCAT(' powered=', BOOL_TO_STRING(bPowered)));
State := CONCAT(State, CONCAT(' unlock=', BOOL_TO_STRING(fb.bUnlock)));
State := CONCAT(State, CONCAT(' unlocked=', BOOL_TO_STRING(fb.bUnlocked)));
State := CONCAT(State, CONCAT(' timeout=', BOOL_TO_STRING(fb.bPowerTimeout)));
State := CONCAT(State, CONCAT(' starts=', INT_TO_STRING(nStarts)));
END_METHOD

END_FUNCTION_BLOCK

// ---- POUs/FB_BrakeCloseHold_Tests.TcPOU
// HalfBROT.FB_BrakeCloseHold (MONETcommon#277): the NC enable of a moving, enabled axis is kept when the brake gate closes under
// it, for its stop; never a new enable against a closed brake, never for a disabled axis, never at standstill, at most tMaxHold.
// The block is called several times per test, one call per PLC cycle it models. Times are T#0S ("no hold"), T#1H ("never within
// a test") or, in the one multi-cycle test, 100 ms of real time.
FUNCTION_BLOCK FB_BrakeCloseHold_Tests EXTENDS TcUnit.FB_TestSuite
VAR
END_VAR

Gate_Closes_Under_Motion_Keeps_Enable();
Closed_Brake_Never_Enables();
Disabled_Axis_Is_Not_Held();
Standstill_Is_Not_Held();
Hold_Ends_At_Standstill_And_Stays_Off();
Gate_Opening_Ends_The_Hold();
Disable_During_Hold_Drops_At_Once();
Zero_Hold_Time_Is_The_Old_Behaviour();
Hold_Ends_After_Max_Time();

// Enabled through the gate and moving, then the gate closes (the shared brake closed): the enable stays on, bHolding is set.
METHOD PRIVATE Gate_Closes_Under_Motion_Keeps_Enable
VAR
	fb	: HalfBROT.FB_BrakeCloseHold;
END_VAR
TEST('Gate_Closes_Under_Motion_Keeps_Enable');
fb(bEnable := TRUE, bBrakeEnable := TRUE, bMoving := TRUE, tMaxHold := T#1H);
AssertTrue(Condition := fb.bAxisEnable, Message := 'enabled through the gate');
AssertFalse(Condition := fb.bHolding, Message := 'no hold while the gate is open');
fb(bEnable := TRUE, bBrakeEnable := FALSE, bMoving := TRUE, tMaxHold := T#1H);
AssertTrue(Condition := fb.bAxisEnable, Message := 'enable kept after the gate closed');
AssertTrue(Condition := fb.bHolding, Message := 'holding');
fb(bEnable := TRUE, bBrakeEnable := FALSE, bMoving := TRUE, tMaxHold := T#1H);
AssertTrue(Condition := fb.bAxisEnable, Message := 'still kept in the next cycle');
TEST_FINISHED();
END_METHOD

// An axis that was not enabled is not enabled against a closed brake, even if it is wanted and reported moving.
METHOD PRIVATE Closed_Brake_Never_Enables
VAR
	fb	: HalfBROT.FB_BrakeCloseHold;
END_VAR
TEST('Closed_Brake_Never_Enables');
fb(bEnable := TRUE, bBrakeEnable := FALSE, bMoving := TRUE, tMaxHold := T#1H);
AssertFalse(Condition := fb.bAxisEnable, Message := 'first cycle: not enabled');
fb(bEnable := TRUE, bBrakeEnable := FALSE, bMoving := TRUE, tMaxHold := T#1H);
AssertFalse(Condition := fb.bAxisEnable, Message := 'second cycle: not enabled');
AssertFalse(Condition := fb.bHolding, Message := 'no hold');
TEST_FINISHED();
END_METHOD

// The controller disables the axis (the faulty one) in the cycle the gate closes: the enable drops at once.
METHOD PRIVATE Disabled_Axis_Is_Not_Held
VAR
	fb	: HalfBROT.FB_BrakeCloseHold;
END_VAR
TEST('Disabled_Axis_Is_Not_Held');
fb(bEnable := TRUE, bBrakeEnable := TRUE, bMoving := TRUE, tMaxHold := T#1H);
fb(bEnable := FALSE, bBrakeEnable := FALSE, bMoving := TRUE, tMaxHold := T#1H);
AssertFalse(Condition := fb.bAxisEnable, Message := 'not enabled');
AssertFalse(Condition := fb.bHolding, Message := 'no hold');
TEST_FINISHED();
END_METHOD

// The gate closes under an axis at standstill (a normal park, a pressure loss at rest): the enable drops at once, as before.
METHOD PRIVATE Standstill_Is_Not_Held
VAR
	fb	: HalfBROT.FB_BrakeCloseHold;
END_VAR
TEST('Standstill_Is_Not_Held');
fb(bEnable := TRUE, bBrakeEnable := TRUE, bMoving := FALSE, tMaxHold := T#1H);
fb(bEnable := TRUE, bBrakeEnable := FALSE, bMoving := FALSE, tMaxHold := T#1H);
AssertFalse(Condition := fb.bAxisEnable, Message := 'not enabled');
AssertFalse(Condition := fb.bHolding, Message := 'no hold');
TEST_FINISHED();
END_METHOD

// The held axis comes to rest: the enable drops, and a later motion report does not bring it back while the gate is closed.
METHOD PRIVATE Hold_Ends_At_Standstill_And_Stays_Off
VAR
	fb	: HalfBROT.FB_BrakeCloseHold;
END_VAR
TEST('Hold_Ends_At_Standstill_And_Stays_Off');
fb(bEnable := TRUE, bBrakeEnable := TRUE, bMoving := TRUE, tMaxHold := T#1H);
fb(bEnable := TRUE, bBrakeEnable := FALSE, bMoving := TRUE, tMaxHold := T#1H);
AssertTrue(Condition := fb.bHolding, Message := 'holding');
fb(bEnable := TRUE, bBrakeEnable := FALSE, bMoving := FALSE, tMaxHold := T#1H);
AssertFalse(Condition := fb.bAxisEnable, Message := 'enable dropped at standstill');
AssertFalse(Condition := fb.bHolding, Message := 'hold ended');
fb(bEnable := TRUE, bBrakeEnable := FALSE, bMoving := TRUE, tMaxHold := T#1H);
AssertFalse(Condition := fb.bAxisEnable, Message := 'no new hold against the closed brake');
TEST_FINISHED();
END_METHOD

// The brake opens again during the hold: the gate takes over, bHolding is cleared, the enable stays on.
METHOD PRIVATE Gate_Opening_Ends_The_Hold
VAR
	fb	: HalfBROT.FB_BrakeCloseHold;
END_VAR
TEST('Gate_Opening_Ends_The_Hold');
fb(bEnable := TRUE, bBrakeEnable := TRUE, bMoving := TRUE, tMaxHold := T#1H);
fb(bEnable := TRUE, bBrakeEnable := FALSE, bMoving := TRUE, tMaxHold := T#1H);
fb(bEnable := TRUE, bBrakeEnable := TRUE, bMoving := TRUE, tMaxHold := T#1H);
AssertTrue(Condition := fb.bAxisEnable, Message := 'enabled through the gate');
AssertFalse(Condition := fb.bHolding, Message := 'hold ended');
TEST_FINISHED();
END_METHOD

// The controller disables the held axis (its stop is over, or another error): the enable drops in the same cycle.
METHOD PRIVATE Disable_During_Hold_Drops_At_Once
VAR
	fb	: HalfBROT.FB_BrakeCloseHold;
END_VAR
TEST('Disable_During_Hold_Drops_At_Once');
fb(bEnable := TRUE, bBrakeEnable := TRUE, bMoving := TRUE, tMaxHold := T#1H);
fb(bEnable := TRUE, bBrakeEnable := FALSE, bMoving := TRUE, tMaxHold := T#1H);
fb(bEnable := FALSE, bBrakeEnable := FALSE, bMoving := TRUE, tMaxHold := T#1H);
AssertFalse(Condition := fb.bAxisEnable, Message := 'enable dropped');
AssertFalse(Condition := fb.bHolding, Message := 'hold ended');
TEST_FINISHED();
END_METHOD

// tMaxHold = T#0S: the enable follows the gate, as before #277.
METHOD PRIVATE Zero_Hold_Time_Is_The_Old_Behaviour
VAR
	fb	: HalfBROT.FB_BrakeCloseHold;
END_VAR
TEST('Zero_Hold_Time_Is_The_Old_Behaviour');
fb(bEnable := TRUE, bBrakeEnable := TRUE, bMoving := TRUE, tMaxHold := T#0S);
AssertTrue(Condition := fb.bAxisEnable, Message := 'enabled through the gate');
fb(bEnable := TRUE, bBrakeEnable := FALSE, bMoving := TRUE, tMaxHold := T#0S);
AssertFalse(Condition := fb.bAxisEnable, Message := 'enable dropped with the gate');
AssertFalse(Condition := fb.bHolding, Message := 'no hold');
TEST_FINISHED();
END_METHOD

// A held axis that never reports standstill: the enable drops after tMaxHold (100 ms, real time; the test gives up after 2 s)
// and does not come back. Multi-cycle: one call per PLC cycle, asserted once at the end.
METHOD PRIVATE Hold_Ends_After_Max_Time
VAR_INST
	fb			: HalfBROT.FB_BrakeCloseHold;
	nStep		: INT;
	tonLimit	: TON;
	tonEarly	: TON;
	bDroppedEarly	: BOOL;
END_VAR
IF nStep >= 99 THEN
	RETURN;
END_IF
TEST('Hold_Ends_After_Max_Time');
CASE nStep OF
0:
	fb(bEnable := TRUE, bBrakeEnable := TRUE, bMoving := TRUE, tMaxHold := T#100MS);
	fb(bEnable := TRUE, bBrakeEnable := FALSE, bMoving := TRUE, tMaxHold := T#100MS);
	nStep := 10;
10:
	fb(bEnable := TRUE, bBrakeEnable := FALSE, bMoving := TRUE, tMaxHold := T#100MS);
	tonLimit(IN := TRUE, PT := T#2S);
	tonEarly(IN := TRUE, PT := T#50MS);
	IF NOT fb.bAxisEnable AND NOT tonEarly.Q THEN
		bDroppedEarly := TRUE;
	END_IF
	IF NOT fb.bAxisEnable OR tonLimit.Q THEN
		fb(bEnable := TRUE, bBrakeEnable := FALSE, bMoving := TRUE, tMaxHold := T#100MS);
		AssertFalse(Condition := fb.bAxisEnable, Message := 'enable dropped after tMaxHold and stays off');
		AssertFalse(Condition := bDroppedEarly, Message := 'not dropped within the first 50 ms');
		AssertFalse(Condition := fb.bHolding, Message := 'hold ended');
		nStep := 99;
		TEST_FINISHED();
	END_IF
END_CASE
END_METHOD

END_FUNCTION_BLOCK

// ---- POUs/F_FocusHoldOnStop_Tests.TcPOU
// HalfBROT.F_FocusHoldOnStop (MONETcommon#278): the hold of FB_FocusControl.Stop() takes the actual position only while the target
// is still the one of the Stop(); a new target set during the stop is kept.
FUNCTION_BLOCK F_FocusHoldOnStop_Tests EXTENDS TcUnit.FB_TestSuite
VAR
END_VAR

Unchanged_Target_Is_Held();
Change_Within_Tolerance_Is_Held();
New_Target_After_Stop_Is_Kept();
Uncalibrated_Focus_Is_Not_Held();

METHOD PRIVATE Unchanged_Target_Is_Held
TEST('Unchanged_Target_Is_Held');
AssertTrue(Condition := HalfBROT.F_FocusHoldOnStop(bCalibrated := TRUE, fTarget := 53.7786, fStopTarget := 53.7786, fTolerance := 0.005),
	Message := 'the target of the Stop(): hold the position reached');
TEST_FINISHED();
END_METHOD

METHOD PRIVATE Change_Within_Tolerance_Is_Held
TEST('Change_Within_Tolerance_Is_Held');
AssertTrue(Condition := HalfBROT.F_FocusHoldOnStop(bCalibrated := TRUE, fTarget := 53.782, fStopTarget := 53.7786, fTolerance := 0.005),
	Message := 'within the tolerance it is the same target');
TEST_FINISHED();
END_METHOD

// MONET/N 2026-11-13 run A of MONETcommon#277: the park sets the focus park position right after the stop of the ramp.
METHOD PRIVATE New_Target_After_Stop_Is_Kept
TEST('New_Target_After_Stop_Is_Kept');
AssertFalse(Condition := HalfBROT.F_FocusHoldOnStop(bCalibrated := TRUE, fTarget := 50.0, fStopTarget := 53.7786, fTolerance := 0.005),
	Message := 'a target set after the Stop() is not overwritten');
TEST_FINISHED();
END_METHOD

METHOD PRIVATE Uncalibrated_Focus_Is_Not_Held
TEST('Uncalibrated_Focus_Is_Not_Held');
AssertFalse(Condition := HalfBROT.F_FocusHoldOnStop(bCalibrated := FALSE, fTarget := 53.7786, fStopTarget := 53.7786, fTolerance := 0.005),
	Message := 'an uncalibrated position is not a target');
TEST_FINISHED();
END_METHOD

END_FUNCTION_BLOCK
